(* IEC 61131-3 sources: ZPLC/conformance/cmp, 592 files *)

(* ---- cmp-042-type-from-another-file-in-a-structure-point.st ---- *)
TYPE Point : STRUCT
  x : INT;
  y : INT;
END_STRUCT END_TYPE

(* ---- cmp-042-global-in-another-file-globals.st ---- *)
VAR_GLOBAL Shared : INT; END_VAR

(* ---- cmp-042-global-initial-value-is-applied-once-globals.st ---- *)
VAR_GLOBAL
  Counter : INT := 100;
END_VAR

(* ---- cmp-042-two-tasks-share-a-global-globals.st ---- *)
VAR_GLOBAL
  Shared : INT;
END_VAR

(* ---- cmp-042-function-from-another-file-in-two-programs-lib.st ---- *)
FUNCTION Twice : INT
VAR_INPUT x : INT; END_VAR
  Twice := x * 2;
END_FUNCTION

(* ---- cmp-004-user-names-case-insensitive.st ---- *)
TYPE
  Pair : STRUCT
    Low : INT;
    High : INT;
  END_STRUCT
  Mode : (Idle, Busy);
END_TYPE

FUNCTION Twice : INT
VAR_INPUT Amount : INT; END_VAR
  TWICE := amount * 2;
END_FUNCTION

FUNCTION_BLOCK Counter
VAR_INPUT Step : INT; END_VAR
VAR_OUTPUT Total : INT; END_VAR
  total := TOTAL + step;
END_FUNCTION_BLOCK

PROGRAM Names
VAR
  P : Pair;
  C : counter;
  M : mode;
  result AT %QW0 : INT;
  is_busy AT %QX2.0 : BOOL;
END_VAR
  p.LOW := twice(AMOUNT := 3);
  p.high := TWICE(4);
  C(STEP := 5);
  c(step := 6);
  M := BUSY;
  result := P.low + p.HIGH + c.TOTAL;
  is_busy := m = busy;
END_PROGRAM

(* ---- cmp-006-missing-base-block.st ---- *)
FUNCTION_BLOCK Child EXTENDS Parent
END_FUNCTION_BLOCK

PROGRAM Caller
VAR
  c : Child;
END_VAR
END_PROGRAM

(* ---- cmp-006-property-is-rejected.st ---- *)
FUNCTION_BLOCK Holder
VAR
  stored : INT;
END_VAR
PROPERTY Value : INT
GET
  Value := stored;
END_GET
END_PROPERTY
END_FUNCTION_BLOCK

PROGRAM Props
VAR
  q AT %QW0 : INT;
END_VAR
  q := 1;
END_PROGRAM

(* ---- cmp-006-unknown-identifier-in-block-body.st ---- *)
FUNCTION_BLOCK Scale
VAR_INPUT a : INT; END_VAR
VAR_OUTPUT b : INT; END_VAR
  b := a * factor;
END_FUNCTION_BLOCK

PROGRAM Caller
VAR
  s : Scale;
  seen AT %QW0 : INT;
END_VAR
  s(a := 2);
  seen := s.b;
END_PROGRAM

(* ---- cmp-006-unknown-member-position.st ---- *)
FUNCTION_BLOCK Counter
VAR_INPUT inc : INT; END_VAR
VAR_OUTPUT total : INT; END_VAR
  total := total + inc;
END_FUNCTION_BLOCK

PROGRAM Typo
VAR
  c : Counter;
END_VAR
  c(nope := 2);
END_PROGRAM

(* ---- cmp-013-int-to-real-in-method-argument.st ---- *)
FUNCTION_BLOCK Scaler
METHOD PUBLIC Twice : REAL
VAR_INPUT
  x : REAL;
END_VAR
  Twice := x * 2.0;
END_METHOD
END_FUNCTION_BLOCK

PROGRAM Caller
VAR
  s : Scaler;
  n : INT := -3;
  r AT %QD0 : REAL;
END_VAR
  r := s.Twice(n);
END_PROGRAM

(* ---- cmp-015-interface-references-stay-one-cell-beside-64-bit-values.st ---- *)
INTERFACE IMeter
METHOD Reading : LREAL
END_METHOD
END_INTERFACE

FUNCTION_BLOCK Probe IMPLEMENTS IMeter
VAR_INPUT
  gain : LREAL;
END_VAR
METHOD Reading : LREAL
  Reading := gain + 0.5;
END_METHOD
END_FUNCTION_BLOCK

FUNCTION_BLOCK Slot
VAR_INPUT
  before : LREAL;
  meter : IMeter;
  after : LINT;
END_VAR
END_FUNCTION_BLOCK

FUNCTION Scaled : LREAL
VAR_INPUT
  source : IMeter;
  factor : LREAL;
  offset : LINT;
END_VAR
  Scaled := source.Reading() * factor + offset;
END_FUNCTION

PROGRAM WideAndInterface
VAR
  a : Probe;
  b : Probe;
  slot : Slot;
  meters : ARRAY[0..1] OF IMeter;
  wide : ARRAY[0..1] OF LINT;
  o_before AT %QD0 : LREAL;
  o_after AT %QD2 : LINT;
  o_slot AT %QD4 : LREAL;
  o_first AT %QD6 : LREAL;
  o_second AT %QD8 : LREAL;
  o_scaled AT %QD10 : LREAL;
  o_wide1 AT %QD12 : LINT;
END_VAR
  a.gain := 1.0;
  b.gain := 2.0;
  slot.before := 1.25;
  slot.meter := b;
  slot.after := -7000000000;
  meters[0] := a;
  meters[1] := b;
  wide[0] := 4294967296;
  wide[1] := -4294967296;
  o_before := slot.before;
  o_after := slot.after;
  o_slot := slot.meter.Reading();
  o_first := meters[0].Reading();
  o_second := meters[1].Reading();
  o_scaled := Scaled(meters[1], 0.1, 3000000000);
  o_wide1 := wide[1];
END_PROGRAM

(* ---- cmp-015-lreal-and-lint-keep-their-place-between-narrow-neighbours.st ---- *)
TYPE Cell :
STRUCT
  flag : BOOL;
  value : LREAL;
  tag : BYTE;
  count : LINT;
  small : INT;
END_STRUCT
END_TYPE

FUNCTION_BLOCK Holder
VAR_INPUT
  on : BOOL;
  level : LREAL;
END_VAR
VAR_OUTPUT
  seen : LINT;
  half : LREAL;
END_VAR
VAR
  steps : BYTE;
END_VAR
  steps := steps + 1;
  seen := seen + 4294967297;
  half := level / 2.0;
END_FUNCTION_BLOCK

PROGRAM WideLayout
VAR
  flag0 : BOOL;
  lone : LREAL;
  byte0 : BYTE;
  wide0 : LINT;
  int0 : INT;
  cells : ARRAY[0..2] OF Cell;
  holder : Holder;
  unit : LINT := 4294967296;
  i : DINT;
  o_flag0 AT %QX512.0 : BOOL;
  o_lone AT %QD0 : LREAL;
  o_byte0 AT %QB1024 : BYTE;
  o_wide0 AT %QD2 : LINT;
  o_int0 AT %QW600 : INT;
  o_flag1 AT %QX512.1 : BOOL;
  o_flag2 AT %QX512.2 : BOOL;
  o_value1 AT %QD4 : LREAL;
  o_value2 AT %QD6 : LREAL;
  o_tag2 AT %QB1025 : BYTE;
  o_count1 AT %QD8 : LINT;
  o_count2 AT %QD10 : LINT;
  o_small1 AT %QW601 : INT;
  o_seen AT %QD12 : LINT;
  o_half AT %QD14 : LREAL;
END_VAR
  flag0 := TRUE;
  lone := 0.1;
  byte0 := 200;
  wide0 := -4294967297;
  int0 := -3;
  FOR i := 0 TO 2 DO
    cells[i].flag := (i = 1);
    cells[i].value := 1.5 * (i + 1);
    cells[i].tag := 10 + i;
    cells[i].count := unit * (i + 1);
    cells[i].small := -100 * (i + 1);
  END_FOR;
  holder(on := TRUE, level := 0.5);
  holder(on := FALSE, level := 0.1);
  o_flag0 := flag0;
  o_lone := lone;
  o_byte0 := byte0;
  o_wide0 := wide0;
  o_int0 := int0;
  o_flag1 := cells[1].flag;
  o_flag2 := cells[2].flag;
  o_value1 := cells[1].value;
  o_value2 := cells[2].value;
  o_tag2 := cells[2].tag;
  o_count1 := cells[1].count;
  o_count2 := cells[2].count;
  o_small1 := cells[1].small;
  o_seen := holder.seen;
  o_half := holder.half;
END_PROGRAM

(* ---- cmp-015-lreal-and-lint-results-of-methods-and-interface-calls.st ---- *)
INTERFACE IMeter
METHOD Reading : LREAL
END_METHOD
METHOD Ticks : LINT
END_METHOD
END_INTERFACE

FUNCTION_BLOCK Probe IMPLEMENTS IMeter
VAR_INPUT
  gain : LREAL;
  offset : LINT;
END_VAR
METHOD Reading : LREAL
  Reading := gain * 0.1 + 0.5;
END_METHOD
METHOD Ticks : LINT
  Ticks := offset * 3;
END_METHOD
METHOD Twice : LREAL
  Twice := Reading() * 2.0;
END_METHOD
END_FUNCTION_BLOCK

FUNCTION_BLOCK FineProbe EXTENDS Probe
METHOD OVERRIDE Reading : LREAL
  Reading := SUPER^.Reading() + 0.25;
END_METHOD
METHOD OVERRIDE Ticks : LINT
  Ticks := SUPER^.Ticks() + 4294967296;
END_METHOD
END_FUNCTION_BLOCK

PROGRAM WideMethods
VAR
  plain : Probe;
  fine : FineProbe;
  meter : IMeter;
  o_reading AT %QD0 : LREAL;
  o_ticks AT %QD2 : LINT;
  o_twice AT %QD4 : LREAL;
  o_fine AT %QD6 : LREAL;
  o_fine_ticks AT %QD8 : LINT;
  o_fine_twice AT %QD10 : LREAL;
  o_through AT %QD12 : LREAL;
  o_through_ticks AT %QD14 : LINT;
  o_through_plain AT %QD16 : LREAL;
  o_after AT %QX512.0 : BOOL;
END_VAR
  plain.gain := 3.0;
  plain.offset := -2000000000;
  fine.gain := 3.0;
  fine.offset := 1;
  o_reading := plain.Reading();
  o_ticks := plain.Ticks();
  o_twice := plain.Twice();
  o_fine := fine.Reading();
  o_fine_ticks := fine.Ticks();
  o_fine_twice := fine.Twice();
  meter := fine;
  o_through := meter.Reading() + 1.0;
  o_through_ticks := meter.Ticks() - 1;
  meter := plain;
  o_through_plain := meter.Reading();
  o_after := meter.Ticks() < 0;
END_PROGRAM

(* ---- cmp-015-lreal-and-lint-through-references-and-in-out-parameters.st ---- *)
FUNCTION_BLOCK Accumulate
VAR_IN_OUT
  total : LREAL;
  count : LINT;
END_VAR
VAR_INPUT
  step : LREAL;
END_VAR
  total := total + step;
  count := count + 1;
END_FUNCTION_BLOCK

PROGRAM WideReferences
VAR
  sum : LREAL;
  big : LINT := 5000000000;
  pd : REF_TO LREAL;
  pl : REF_TO LINT;
  acc : Accumulate;
  n : LINT;
  o_sum AT %QD0 : LREAL;
  o_big AT %QD2 : LINT;
  o_count AT %QD4 : LINT;
  o_through AT %QD6 : LREAL;
END_VAR
  pd := REF(sum);
  pl := REF(big);
  acc(total := sum, count := n, step := 0.5);
  acc(total := sum, count := n, step := 0.25);
  pd^ := pd^ + 1.0;
  pl^ := pl^ * 2;
  o_sum := sum;
  o_big := big;
  o_count := n;
  o_through := pd^ * 2.0;
END_PROGRAM

(* ---- cmp-019-fb-member-int.st ---- *)
FUNCTION_BLOCK Big
VAR_OUTPUT o : INT; END_VAR
  o := 1000;
END_FUNCTION_BLOCK

PROGRAM Member
VAR
  f : Big;
  seen AT %QW0 : INT;
END_VAR
  f();
  seen := f.o;
END_PROGRAM

(* ---- cmp-019-fb-mixed-width-members.st ---- *)
FUNCTION_BLOCK Mixed
VAR_INPUT b : BYTE; END_VAR
VAR_OUTPUT i : INT; d : DINT; r : REAL; s : SINT; END_VAR
  i := -1000;
  d := -100000;
  r := 2.5;
  s := -3;
  b := 200;
END_FUNCTION_BLOCK

PROGRAM Main
VAR
  m : Mixed;
  oi AT %QW0 : INT;
  od AT %QD1 : DINT;
  orr AT %QD2 : REAL;
  os AT %QB12 : SINT;
  ob AT %QB13 : BYTE;
END_VAR
  m();
  oi := m.i;
  od := m.d;
  orr := m.r;
  os := m.s;
  ob := m.b;
END_PROGRAM

(* ---- cmp-021-fb-string-member-initial-value.st ---- *)
FUNCTION_BLOCK Named
VAR_OUTPUT label : STRING[16] := 'unit'; END_VAR
END_FUNCTION_BLOCK

PROGRAM Main
VAR
  n : Named;
  l AT %QW0 : INT;
  ok AT %QX2.0 : BOOL;
END_VAR
  n();
  l := LEN(n.label);
  ok := n.label = 'unit';
END_PROGRAM

(* ---- cmp-024-null-inside-a-function-block.st ---- *)
FUNCTION_BLOCK Probe
VAR_INPUT bind : BOOL; target : DINT; END_VAR
VAR_OUTPUT isNull : BOOL; value : DINT; END_VAR
VAR p : REF_TO DINT; END_VAR
  IF bind THEN
    p := REF(target);
  ELSE
    p := NULL;
  END_IF;
  isNull := p = NULL;
  IF NOT isNull THEN
    value := p^;
  END_IF;
END_FUNCTION_BLOCK

PROGRAM Main
VAR
  probe : Probe;
  a AT %QX0.0 : BOOL;
  b AT %QX0.1 : BOOL;
  v AT %QD1 : DINT;
END_VAR
  probe(bind := FALSE, target := 5);
  a := probe.isNull;
  probe(bind := TRUE, target := 123456);
  b := probe.isNull;
  v := probe.value;
END_PROGRAM

(* ---- cmp-025-fb-instances-keep-their-own-initial-values.st ---- *)
FUNCTION_BLOCK Start
VAR_OUTPUT v : INT := 5; END_VAR
  v := v + 1;
END_FUNCTION_BLOCK

PROGRAM Main
VAR
  f1 : Start := (v := 10);
  f2 : Start;
  a AT %QW0 : INT;
  b AT %QW1 : INT;
END_VAR
  f1();
  f2();
  a := f1.v;
  b := f2.v;
END_PROGRAM

(* ---- cmp-025-fb-member-initial-value.st ---- *)
FUNCTION_BLOCK Start
VAR_OUTPUT v : INT := 5; END_VAR
  v := v + 1;
END_FUNCTION_BLOCK

PROGRAM Members
VAR
  f : Start;
  seen AT %QW0 : INT;
END_VAR
  f();
  seen := f.v;
END_PROGRAM

(* ---- cmp-025-var-input-and-var-output-of-a-function-block.st ---- *)
FUNCTION_BLOCK Accumulate
VAR_INPUT step : INT; END_VAR
VAR_OUTPUT total : INT; END_VAR
  total := total + step;
END_FUNCTION_BLOCK

PROGRAM Inputs
VAR
  acc : Accumulate;
  result AT %QW0 : INT;
END_VAR
  acc(step := 3);
  result := acc.total;
END_PROGRAM

(* ---- cmp-026-function-block-constant-assignment-rejected.st ---- *)
FUNCTION_BLOCK Limit
VAR_OUTPUT clipped : INT; END_VAR
VAR CONSTANT MAXV : INT := 100; END_VAR
  MAXV := 5;
  clipped := MAXV;
END_FUNCTION_BLOCK

PROGRAM Main
VAR
  l : Limit;
END_VAR
  l();
END_PROGRAM

(* ---- cmp-026-function-block-constant-member.st ---- *)
FUNCTION_BLOCK Limit
VAR_INPUT v : INT; END_VAR
VAR_OUTPUT clipped : INT; END_VAR
VAR CONSTANT MAXV : INT := 100; END_VAR
  IF v > MAXV THEN
    clipped := MAXV;
  ELSE
    clipped := v;
  END_IF;
END_FUNCTION_BLOCK

PROGRAM Main
VAR
  l : Limit;
  out AT %QW0 : INT;
END_VAR
  l(v := 250);
  out := l.clipped;
END_PROGRAM

(* ---- cmp-027-fb-var-temp-initial-value-on-every-call.st ---- *)
FUNCTION_BLOCK Temp
VAR_OUTPUT o : INT; END_VAR
VAR_TEMP k : INT := 10; END_VAR
  k := k + 1;
  o := k;
END_FUNCTION_BLOCK

PROGRAM Main
VAR
  f : Temp;
  seen AT %QW0 : INT;
END_VAR
  f();
  seen := f.o;
END_PROGRAM

(* ---- cmp-027-fb-var-temp-not-retained.st ---- *)
FUNCTION_BLOCK Temp
VAR_OUTPUT o : INT; END_VAR
VAR_TEMP k : INT; END_VAR
  k := k + 1;
  o := k;
END_FUNCTION_BLOCK

PROGRAM Calls
VAR
  f : Temp;
  seen AT %QW0 : INT;
END_VAR
  f();
  seen := f.o;
END_PROGRAM

(* ---- cmp-028-in-out-bound-to-member-and-element.st ---- *)
TYPE Pt : STRUCT x : INT; z : DINT; END_STRUCT END_TYPE

FUNCTION_BLOCK Inc
VAR_IN_OUT x : INT; END_VAR
  x := x + 1;
END_FUNCTION_BLOCK

PROGRAM Main
VAR
  f : Inc;
  s : Pt;
  a : ARRAY[0..3] OF INT;
  i : INT;
  sx AT %QW0 : INT;
  a2 AT %QW1 : INT;
  a1 AT %QW2 : INT;
END_VAR
  s.x := 40;
  i := 2;
  a[2] := 7;
  f(x := s.x);
  f(x := a[i]);
  sx := s.x;
  a2 := a[2];
  a1 := a[1];
END_PROGRAM

(* ---- cmp-028-in-out-of-another-type-rejected.st ---- *)
FUNCTION_BLOCK Inc
VAR_IN_OUT x : INT; END_VAR
  x := x + 1;
END_FUNCTION_BLOCK

PROGRAM Main
VAR
  f : Inc;
  d : DINT;
END_VAR
  f(x := d);
END_PROGRAM

(* ---- cmp-028-in-out-two-instances-different-targets.st ---- *)
FUNCTION_BLOCK Inc
VAR_IN_OUT x : DINT; END_VAR
  x := x + 100000;
END_FUNCTION_BLOCK

PROGRAM Main
VAR
  f : Inc;
  g : Inc;
  a : DINT := 1;
  b : DINT := 2;
  oa AT %QD0 : DINT;
  ob AT %QD1 : DINT;
END_VAR
  f(x := a);
  g(x := b);
  f();
  oa := a;
  ob := b;
END_PROGRAM

(* ---- cmp-028-in-out-whole-structure.st ---- *)
TYPE Pt : STRUCT x : INT; z : DINT; END_STRUCT END_TYPE

FUNCTION_BLOCK Move
VAR_IN_OUT p : Pt; END_VAR
  p.x := p.x + 1;
  p.z := p.z + 100000;
END_FUNCTION_BLOCK

PROGRAM Main
VAR
  m : Move;
  point : Pt;
  ox AT %QW0 : INT;
  oz AT %QD1 : DINT;
END_VAR
  point.x := 5;
  point.z := 1;
  m(p := point);
  ox := point.x;
  oz := point.z;
END_PROGRAM

(* ---- cmp-028-unbound-in-out-faults.st ---- *)
FUNCTION_BLOCK Inc
VAR_IN_OUT x : INT; END_VAR
  x := x + 1;
END_FUNCTION_BLOCK

PROGRAM Main
VAR
  f : Inc;
END_VAR
  f();
END_PROGRAM

(* ---- cmp-028-var-in-out-by-reference.st ---- *)
FUNCTION_BLOCK Inc
VAR_IN_OUT x : INT; END_VAR
  x := x + 1;
END_FUNCTION_BLOCK

PROGRAM Reference
VAR
  f : Inc;
  v : INT := 5;
  seen AT %QW0 : INT;
END_VAR
  f(x := v);
  seen := v;
END_PROGRAM

(* ---- cmp-030-var-external-in-function-block.st ---- *)
VAR_GLOBAL
  hits : INT;
END_VAR

FUNCTION_BLOCK Counter
VAR_EXTERNAL hits : INT; END_VAR
  hits := hits + 1;
END_FUNCTION_BLOCK

PROGRAM Shared
VAR
  a : Counter;
  b : Counter;
  seen AT %QW0 : INT;
END_VAR
  a();
  b();
  seen := hits;
END_PROGRAM

(* ---- cmp-033-library-names-as-names-of-everything.st ---- *)
TYPE Reading : STRUCT Pulse : INT; Blink : INT; END_STRUCT END_TYPE

FUNCTION_BLOCK Scale
VAR_INPUT Counter : INT; END_VAR
VAR_OUTPUT Pwm : INT; END_VAR
  Pwm := Counter * 2;
END_FUNCTION_BLOCK

FUNCTION Twice : INT
VAR_INPUT Ton : INT; END_VAR
  Twice := Ton + Ton;
END_FUNCTION

PROGRAM Names
VAR
  Fifo : Reading;
  Lifo : Scale;
  Rs : INT;
  sum AT %QW0 : INT;
END_VAR
  Fifo.Pulse := 3;
  Fifo.Blink := 4;
  Lifo(Counter := Fifo.Pulse);
  Rs := Twice(Ton := Fifo.Blink);
  sum := Lifo.Pwm + Rs;
END_PROGRAM

(* ---- cmp-033-user-block-named-like-a-library-block.st ---- *)
FUNCTION_BLOCK Blink
VAR_OUTPUT level : INT; END_VAR
  level := 7;
END_FUNCTION_BLOCK

PROGRAM Own
VAR
  b : blink;
  seen AT %QW0 : INT;
END_VAR
  b();
  seen := b.level;
END_PROGRAM

(* ---- cmp-036-return-leaves-the-function-block-only.st ---- *)
FUNCTION_BLOCK Gate
VAR_INPUT go : BOOL; END_VAR
VAR_OUTPUT q : INT; END_VAR
  q := 1;
  IF go THEN
    q := 5;
    RETURN;
  END_IF;
  q := 9;
END_FUNCTION_BLOCK

PROGRAM Returns
VAR
  g : Gate;
  early AT %QW0 : INT;
  after AT %QX2.0 : BOOL;
END_VAR
  g(go := TRUE);
  early := g.q;
  after := TRUE;
END_PROGRAM

(* ---- cmp-037-output-assigned-with-colon-equals-is-rejected.st ---- *)
FUNCTION_BLOCK Adder
VAR_INPUT a : INT; END_VAR
VAR_OUTPUT sum : INT; END_VAR
  sum := a;
END_FUNCTION_BLOCK

PROGRAM Binding
VAR
  add : Adder;
END_VAR
  add(a := 1, sum := 2);
END_PROGRAM

(* ---- cmp-037-output-binding-of-a-user-block.st ---- *)
FUNCTION_BLOCK Adder
VAR_INPUT a : INT; b : INT; END_VAR
VAR_OUTPUT sum : INT; big : BOOL; END_VAR
  sum := a + b;
  big := sum > 100;
END_FUNCTION_BLOCK

PROGRAM Binding
VAR
  add : Adder;
  total AT %QW0 : INT;
  large AT %QX2.0 : BOOL;
END_VAR
  add(a := 60, b := 70, sum => total, big => large);
END_PROGRAM

(* ---- cmp-037-positional-call-of-a-user-block-is-rejected.st ---- *)
FUNCTION_BLOCK Adder
VAR_INPUT a : INT; END_VAR
VAR_OUTPUT sum : INT; END_VAR
  sum := a;
END_FUNCTION_BLOCK

PROGRAM Binding
VAR
  add : Adder;
END_VAR
  add(1);
END_PROGRAM

(* ---- cmp-037-unknown-parameter-of-a-user-block.st ---- *)
FUNCTION_BLOCK Adder
VAR_INPUT a : INT; END_VAR
VAR_OUTPUT sum : INT; END_VAR
  sum := a;
END_FUNCTION_BLOCK

PROGRAM Binding
VAR
  add : Adder;
END_VAR
  add(a := 1, nothing := 2);
END_PROGRAM

(* ---- cmp-038-array-of-user-blocks.st ---- *)
FUNCTION_BLOCK Total
VAR_INPUT inc : INT; END_VAR
VAR_OUTPUT sum : INT; END_VAR
  sum := sum + inc;
END_FUNCTION_BLOCK

PROGRAM Composition
VAR
  t : ARRAY[0..1] OF Total;
  x AT %QW0 : INT;
  y AT %QW2 : INT;
END_VAR
  t[0](inc := 1);
  t[1](inc := 10);
  x := t[0].sum;
  y := t[1].sum;
END_PROGRAM

(* ---- cmp-038-instance-inside-function-block.st ---- *)
FUNCTION_BLOCK Debounce
VAR_INPUT sig : BOOL; END_VAR
VAR_OUTPUT out : BOOL; END_VAR
VAR tmr : TON; END_VAR
  tmr(IN := sig, PT := T#20ms);
  out := tmr.Q;
END_FUNCTION_BLOCK

PROGRAM Composition
VAR
  d : Debounce;
  settled AT %QX0.0 : BOOL;
END_VAR
  d(sig := TRUE);
  settled := d.out;
END_PROGRAM

(* ---- cmp-038-timer-inside-two-instances.st ---- *)
FUNCTION_BLOCK Delay
VAR_INPUT go : BOOL; END_VAR
VAR_OUTPUT done : BOOL; END_VAR
VAR t : TON; END_VAR
  t(IN := go, PT := T#25ms);
  done := t.Q;
END_FUNCTION_BLOCK

PROGRAM Composition
VAR
  fast : Delay;
  idle : Delay;
  a AT %QX0.0 : BOOL;
  b AT %QX0.1 : BOOL;
END_VAR
  fast(go := TRUE);
  idle(go := FALSE);
  a := fast.done;
  b := idle.done;
END_PROGRAM

(* ---- cmp-038-two-instances-keep-own-state.st ---- *)
FUNCTION_BLOCK Counter
VAR_INPUT inc : INT; END_VAR
VAR_OUTPUT total : INT; END_VAR
  total := total + inc;
END_FUNCTION_BLOCK

PROGRAM Composition
VAR
  a : Counter;
  b : Counter;
  x AT %QW0 : INT;
  y AT %QW1 : INT;
END_VAR
  a(inc := 1);
  b(inc := 10);
  x := a.total;
  y := b.total;
END_PROGRAM

(* ---- cmp-039-for-inside-function-block.st ---- *)
FUNCTION_BLOCK Summer
VAR_OUTPUT s : INT; END_VAR
VAR i : INT; END_VAR
  s := 0;
  FOR i := 1 TO 4 DO
    s := s + i;
  END_FOR;
END_FUNCTION_BLOCK

PROGRAM Loop
VAR
  f : Summer;
  sum AT %QW0 : INT;
END_VAR
  f();
  sum := f.s;
END_PROGRAM

(* ---- cmp-041-abstract-block-cannot-be-instantiated.st ---- *)
FUNCTION_BLOCK ABSTRACT Template
METHOD ABSTRACT Step : INT
END_METHOD
END_FUNCTION_BLOCK

PROGRAM Abstraction
VAR
  t : Template;
END_VAR
END_PROGRAM

(* ---- cmp-041-abstract-method-is-run-by-the-derived-block.st ---- *)
FUNCTION_BLOCK ABSTRACT Template
METHOD ABSTRACT Step : INT
END_METHOD
METHOD Run : INT
  Run := Step() * 2 + 1;
END_METHOD
END_FUNCTION_BLOCK

FUNCTION_BLOCK Seven EXTENDS Template
METHOD OVERRIDE Step : INT
  Step := 7;
END_METHOD
END_FUNCTION_BLOCK

FUNCTION_BLOCK Nine EXTENDS Template
METHOD OVERRIDE Step : INT
  Step := 9;
END_METHOD
END_FUNCTION_BLOCK

PROGRAM Abstraction
VAR
  a : Seven;
  b : Nine;
  x AT %QW0 : INT;
  y AT %QW1 : INT;
END_VAR
  x := a.Run();
  y := b.Run();
END_PROGRAM

(* ---- cmp-041-abstract-method-left-unimplemented-is-rejected.st ---- *)
FUNCTION_BLOCK ABSTRACT Template
METHOD ABSTRACT Step : INT
END_METHOD
END_FUNCTION_BLOCK

FUNCTION_BLOCK Lazy EXTENDS Template
END_FUNCTION_BLOCK

PROGRAM Abstraction
VAR
  l : Lazy;
END_VAR
END_PROGRAM

(* ---- cmp-041-final-block-cannot-be-extended.st ---- *)
FUNCTION_BLOCK FINAL Sealed
END_FUNCTION_BLOCK

FUNCTION_BLOCK Open EXTENDS Sealed
END_FUNCTION_BLOCK

PROGRAM Sealing
END_PROGRAM

(* ---- cmp-041-final-method-cannot-be-overridden.st ---- *)
FUNCTION_BLOCK Base
METHOD FINAL Reading : INT
  Reading := 3;
END_METHOD
END_FUNCTION_BLOCK

FUNCTION_BLOCK Derived EXTENDS Base
METHOD OVERRIDE Reading : INT
  Reading := 4;
END_METHOD
END_FUNCTION_BLOCK

PROGRAM Derivation
VAR
  d : Derived;
  q AT %QW0 : INT;
END_VAR
  q := d.Reading();
END_PROGRAM

(* ---- cmp-041-instance-that-does-not-implement-the-interface-is-rejected.st ---- *)
INTERFACE IRun
METHOD Go : INT
END_METHOD
END_INTERFACE

FUNCTION_BLOCK Plain
METHOD Go : INT
  Go := 1;
END_METHOD
END_FUNCTION_BLOCK

PROGRAM Wrong
VAR
  p : Plain;
  r : IRun;
END_VAR
  r := p;
END_PROGRAM

(* ---- cmp-041-interface-call-of-a-null-reference-faults.st ---- *)
INTERFACE IRun
METHOD Go : INT
END_METHOD
END_INTERFACE

FUNCTION_BLOCK A IMPLEMENTS IRun
METHOD Go : INT
  Go := 1;
END_METHOD
END_FUNCTION_BLOCK

PROGRAM Unassigned
VAR
  a : A;
  r : IRun;
  seen AT %QW0 : INT;
END_VAR
  seen := 5;
  seen := r.Go();
END_PROGRAM

(* ---- cmp-041-interface-dispatch-by-the-instance-assigned.st ---- *)
INTERFACE IShape
METHOD Area : INT
END_METHOD
END_INTERFACE

FUNCTION_BLOCK Square IMPLEMENTS IShape
VAR_INPUT side : INT; END_VAR
METHOD Area : INT
  Area := side * side;
END_METHOD
END_FUNCTION_BLOCK

FUNCTION_BLOCK Rectangle IMPLEMENTS IShape
VAR_INPUT width : INT; height : INT; END_VAR
METHOD Area : INT
  Area := width * height;
END_METHOD
END_FUNCTION_BLOCK

PROGRAM Shapes
VAR
  sq : Square;
  rect : Rectangle;
  shape : IShape;
  first AT %QW0 : INT;
  second AT %QW1 : INT;
  third AT %QW2 : INT;
END_VAR
  sq.side := 4;
  rect.width := 3;
  rect.height := 5;
  shape := sq;
  first := shape.Area();
  shape := rect;
  second := shape.Area();
  sq.side := 7;
  shape := sq;
  third := shape.Area();
END_PROGRAM

(* ---- cmp-041-interface-dispatch.st ---- *)
INTERFACE IRun
METHOD Go : INT
END_METHOD
END_INTERFACE

FUNCTION_BLOCK A IMPLEMENTS IRun
METHOD Go : INT
  Go := 1;
END_METHOD
END_FUNCTION_BLOCK

PROGRAM Dispatch
VAR
  a : A;
  r : IRun;
  seen AT %QW0 : INT;
END_VAR
  r := a;
  seen := r.Go();
END_PROGRAM

(* ---- cmp-041-interface-through-inheritance-and-array-elements.st ---- *)
INTERFACE IStep
METHOD Run : INT
END_METHOD
END_INTERFACE

FUNCTION_BLOCK Base IMPLEMENTS IStep
VAR_INPUT n : INT; END_VAR
METHOD Run : INT
  Run := n;
END_METHOD
END_FUNCTION_BLOCK

FUNCTION_BLOCK Derived EXTENDS Base
METHOD OVERRIDE Run : INT
  Run := SUPER^.Run() + 1000;
END_METHOD
END_FUNCTION_BLOCK

PROGRAM Steps
VAR
  plain : ARRAY[0..2] OF Base;
  special : Derived;
  step : IStep;
  i : INT;
  total AT %QW0 : INT;
  last AT %QW1 : INT;
END_VAR
  plain[0].n := 1;
  plain[1].n := 20;
  plain[2].n := 300;
  special.n := 5;
  total := 0;
  FOR i := 0 TO 2 DO
    step := plain[i];
    total := total + step.Run();
  END_FOR;
  step := special;
  last := step.Run();
END_PROGRAM

(* ---- cmp-041-interface-variable-as-an-argument-of-a-function.st ---- *)
INTERFACE IMeasure
METHOD Read : INT
END_METHOD
END_INTERFACE

FUNCTION_BLOCK Fixed IMPLEMENTS IMeasure
METHOD Read : INT
  Read := 40;
END_METHOD
END_FUNCTION_BLOCK

FUNCTION_BLOCK Counted IMPLEMENTS IMeasure
VAR reads : INT; END_VAR
METHOD Read : INT
  reads := reads + 1;
  Read := reads;
END_METHOD
END_FUNCTION_BLOCK

FUNCTION Twice : INT
VAR_INPUT source : IMeasure; END_VAR
  Twice := source.Read() + source.Read();
END_FUNCTION

PROGRAM Sampling
VAR
  f : Fixed;
  c : Counted;
  a AT %QW0 : INT;
  b AT %QW1 : INT;
END_VAR
  a := Twice(source := f);
  b := Twice(source := c);
END_PROGRAM

(* ---- cmp-041-interface-variable-as-an-input-of-a-block.st ---- *)
INTERFACE IGain
METHOD Apply : INT
VAR_INPUT x : INT; END_VAR
END_METHOD
END_INTERFACE

FUNCTION_BLOCK Doubler IMPLEMENTS IGain
METHOD Apply : INT
VAR_INPUT x : INT; END_VAR
  Apply := x * 2;
END_METHOD
END_FUNCTION_BLOCK

FUNCTION_BLOCK Offsetter IMPLEMENTS IGain
VAR offset : INT := 100; END_VAR
METHOD Apply : INT
VAR_INPUT x : INT; END_VAR
  Apply := x + offset;
END_METHOD
END_FUNCTION_BLOCK

FUNCTION_BLOCK Stage
VAR_INPUT gain : IGain; value : INT; END_VAR
VAR_OUTPUT result : INT; END_VAR
  result := gain.Apply(value);
END_FUNCTION_BLOCK

PROGRAM Pipeline
VAR
  d : Doubler;
  o : Offsetter;
  stage : Stage;
  a AT %QW0 : INT;
  b AT %QW1 : INT;
END_VAR
  stage(gain := d, value := 21);
  a := stage.result;
  stage(gain := o, value := 21);
  b := stage.result;
END_PROGRAM

(* ---- cmp-041-method-results-of-each-type-and-inherited-statement-call.st ---- *)
FUNCTION_BLOCK Base
VAR
  n : INT;
END_VAR
METHOD Flag : BOOL
  Flag := n > 0;
END_METHOD
METHOD Small : SINT
  Small := -5;
END_METHOD
METHOD Ratio : REAL
  Ratio := 2.5;
END_METHOD
METHOD Wide : DINT
  Wide := -70000;
END_METHOD
METHOD Bump
  n := n + 1;
END_METHOD
END_FUNCTION_BLOCK

FUNCTION_BLOCK Derived EXTENDS Base
END_FUNCTION_BLOCK

PROGRAM Results
VAR
  d : Derived;
  i : INT;
  q0 AT %QX0.0 : BOOL;
  q1 AT %QB1 : SINT;
  q2 AT %QD1 : REAL;
  q3 AT %QD2 : DINT;
  q4 AT %QW6 : INT;
END_VAR
  FOR i := 1 TO 20 DO
    d.Flag();
    d.Bump();
  END_FOR;
  q0 := d.Flag();
  q1 := d.Small();
  q2 := d.Ratio();
  q3 := d.Wide();
  q4 := d.n;
END_PROGRAM

(* ---- cmp-041-method-with-several-assignments-called-in-a-loop.st ---- *)
FUNCTION_BLOCK Chooser
VAR
  calls : INT;
END_VAR
METHOD Pick : INT
VAR_INPUT
  x : INT;
END_VAR
  Pick := x;
  IF x > 5 THEN
    Pick := x * 2;
  END_IF;
  IF x > 8 THEN
    Pick := 0 - x;
  END_IF;
  calls := calls + 1;
END_METHOD
METHOD Never : INT
  calls := calls + 100;
END_METHOD
END_FUNCTION_BLOCK

PROGRAM Loop
VAR
  c : Chooser;
  i : INT;
  total : INT;
  nothing : INT := 7;
  q0 AT %QW0 : INT;
  q1 AT %QW1 : INT;
  q2 AT %QW2 : INT;
END_VAR
  total := 0;
  FOR i := 1 TO 10 DO
    total := total + c.Pick(i);
  END_FOR;
  nothing := c.Never();
  c.Pick(3);
  q0 := total;
  q1 := c.calls;
  q2 := nothing;
END_PROGRAM

(* ---- cmp-041-override-and-inherited-method.st ---- *)
FUNCTION_BLOCK Base
METHOD A : INT
  A := 1;
END_METHOD
METHOD B : INT
  B := 10;
END_METHOD
END_FUNCTION_BLOCK

FUNCTION_BLOCK Derived EXTENDS Base
METHOD OVERRIDE B : INT
  B := 20;
END_METHOD
END_FUNCTION_BLOCK

PROGRAM Inheritance
VAR
  d : Derived;
  x AT %QW0 : INT;
  y AT %QW1 : INT;
END_VAR
  x := d.A();
  y := d.B();
END_PROGRAM

(* ---- cmp-041-private-method-is-not-callable-from-a-derived-block.st ---- *)
FUNCTION_BLOCK Sensor
METHOD PRIVATE Offset : INT
  Offset := 2;
END_METHOD
END_FUNCTION_BLOCK

FUNCTION_BLOCK Scaled EXTENDS Sensor
METHOD Shifted : INT
  Shifted := Offset();
END_METHOD
END_FUNCTION_BLOCK

PROGRAM Access
VAR
  s : Scaled;
  a AT %QW0 : INT;
END_VAR
  a := s.Shifted();
END_PROGRAM

(* ---- cmp-041-private-method-is-not-callable-from-outside.st ---- *)
FUNCTION_BLOCK Gauge
METHOD PRIVATE Reading : INT
  Reading := 3;
END_METHOD
END_FUNCTION_BLOCK

PROGRAM Access
VAR
  g : Gauge;
  q AT %QW0 : INT;
END_VAR
  q := g.Reading();
END_PROGRAM

(* ---- cmp-041-protected-method-is-callable-from-a-derived-block.st ---- *)
FUNCTION_BLOCK Sensor
METHOD PROTECTED Raw : INT
  Raw := 21;
END_METHOD
METHOD PRIVATE Offset : INT
  Offset := 2;
END_METHOD
METHOD PUBLIC Corrected : INT
  Corrected := Raw() + Offset();
END_METHOD
END_FUNCTION_BLOCK

FUNCTION_BLOCK Scaled EXTENDS Sensor
METHOD Doubled : INT
  Doubled := Raw() * 2;
END_METHOD
END_FUNCTION_BLOCK

PROGRAM Access
VAR
  s : Scaled;
  a AT %QW0 : INT;
  b AT %QW1 : INT;
END_VAR
  a := s.Corrected();
  b := s.Doubled();
END_PROGRAM

(* ---- cmp-041-protected-method-is-not-callable-from-outside.st ---- *)
FUNCTION_BLOCK Gauge
METHOD PROTECTED Reading : INT
  Reading := 3;
END_METHOD
END_FUNCTION_BLOCK

PROGRAM Access
VAR
  g : Gauge;
  q AT %QW0 : INT;
END_VAR
  q := g.Reading();
END_PROGRAM

(* ---- cmp-041-public-method-is-callable.st ---- *)
FUNCTION_BLOCK Gauge
METHOD PUBLIC Reading : INT
  Reading := 3;
END_METHOD
END_FUNCTION_BLOCK

PROGRAM Access
VAR
  g : Gauge;
  q AT %QW0 : INT;
END_VAR
  q := g.Reading();
END_PROGRAM

(* ---- cmp-041-super-call-of-a-private-method-is-rejected.st ---- *)
FUNCTION_BLOCK Base
METHOD PRIVATE Secret : INT
  Secret := 1;
END_METHOD
END_FUNCTION_BLOCK

FUNCTION_BLOCK Derived EXTENDS Base
METHOD Peek : INT
  Peek := SUPER^.Secret();
END_METHOD
END_FUNCTION_BLOCK

PROGRAM P
VAR
  d : Derived;
  a AT %QW0 : INT;
END_VAR
  a := d.Peek();
END_PROGRAM

(* ---- cmp-041-super-call-runs-the-base-body.st ---- *)
FUNCTION_BLOCK Counter
VAR_OUTPUT total : INT; END_VAR
  total := total + 1;
END_FUNCTION_BLOCK

FUNCTION_BLOCK DoubleCounter EXTENDS Counter
  SUPER^();
  total := total + 10;
END_FUNCTION_BLOCK

PROGRAM Run
VAR
  c : DoubleCounter;
  seen AT %QW0 : INT;
END_VAR
  c();
  c();
  seen := c.total;
END_PROGRAM

(* ---- cmp-041-super-call-through-three-levels.st ---- *)
FUNCTION_BLOCK Base
METHOD Value : INT
  Value := 1;
END_METHOD
END_FUNCTION_BLOCK

FUNCTION_BLOCK Middle EXTENDS Base
METHOD OVERRIDE Value : INT
  Value := SUPER^.Value() + 10;
END_METHOD
END_FUNCTION_BLOCK

FUNCTION_BLOCK Top EXTENDS Middle
METHOD OVERRIDE Value : INT
  Value := SUPER^.Value() + 100;
END_METHOD
END_FUNCTION_BLOCK

PROGRAM Chain
VAR
  t : Top;
  seen AT %QW0 : INT;
END_VAR
  seen := t.Value();
END_PROGRAM

(* ---- cmp-041-super-call.st ---- *)
FUNCTION_BLOCK A
METHOD M : INT
  M := 1;
END_METHOD
END_FUNCTION_BLOCK

FUNCTION_BLOCK B EXTENDS A
METHOD OVERRIDE M : INT
  M := SUPER^.M() + 1;
END_METHOD
END_FUNCTION_BLOCK

PROGRAM Inheritance
VAR
  b : B;
  seen AT %QW0 : INT;
END_VAR
  seen := b.M();
END_PROGRAM

(* ---- cmp-041-this-member-in-method.st ---- *)
FUNCTION_BLOCK Bumper
VAR c : INT; END_VAR
METHOD Bump : INT
  THIS.c := THIS.c + 1;
  Bump := THIS.c;
END_METHOD
END_FUNCTION_BLOCK

PROGRAM Methods
VAR
  m : Bumper;
  seen AT %QW0 : INT;
END_VAR
  seen := m.Bump();
END_PROGRAM

(* ---- cmp-042-debug-map-addresses-of-every-program-lib.st ---- *)
VAR_GLOBAL
  Shared : INT;
END_VAR

FUNCTION_BLOCK Gate
VAR_INPUT open : BOOL; END_VAR
VAR_OUTPUT passed : BOOL; END_VAR
  passed := open;
END_FUNCTION_BLOCK

(* ---- cmp-042-function-block-declared-in-two-files-is-rejected-a.st ---- *)
(* the first declaration *)
FUNCTION_BLOCK Echo
END_FUNCTION_BLOCK

(* ---- cmp-042-function-block-declared-in-two-files-is-rejected-b.st ---- *)
FUNCTION_BLOCK Echo
VAR_INPUT sig : BOOL; END_VAR
END_FUNCTION_BLOCK

(* ---- cmp-042-function-block-in-another-file-echo.st ---- *)
FUNCTION_BLOCK Echo
VAR_INPUT sig : BOOL; END_VAR
VAR_OUTPUT out : BOOL; END_VAR
  out := sig;
END_FUNCTION_BLOCK

(* ---- cmp-001-undeclared-assignment-target.st ---- *)
PROGRAM Typo
VAR
  x : INT;
END_VAR
  nope := 5;
  x := 1;
END_PROGRAM

(* ---- cmp-001-undeclared-identifier-read.st ---- *)
PROGRAM Typo
VAR
  x : INT;
END_VAR
  x := nope + 1;
END_PROGRAM

(* ---- cmp-001-unknown-function.st ---- *)
PROGRAM Typo
VAR
  x : INT;
END_VAR
  x := NOSUCHFN(1);
END_PROGRAM

(* ---- cmp-002-exit-outside-loop.st ---- *)
PROGRAM Typo
VAR
  x : INT;
END_VAR
  EXIT;
  x := 1;
END_PROGRAM

(* ---- cmp-002-wrong-argument-count.st ---- *)
PROGRAM Typo
VAR
  x : INT;
END_VAR
  x := ABS();
END_PROGRAM

(* ---- cmp-003-char-is-rejected.st ---- *)
PROGRAM Character
VAR
  c : CHAR;
  q AT %QW0 : INT;
END_VAR
  q := 1;
END_PROGRAM

(* ---- cmp-003-ldate-is-rejected.st ---- *)
PROGRAM Long
VAR
  d : LDATE;
  q AT %QW0 : INT;
END_VAR
  q := 1;
END_PROGRAM

(* ---- cmp-003-ldt-is-rejected.st ---- *)
PROGRAM Long
VAR
  t : LDT;
  q AT %QW0 : INT;
END_VAR
  q := 1;
END_PROGRAM

(* ---- cmp-003-ltime-is-rejected.st ---- *)
PROGRAM Long
VAR
  t : LTIME;
  q AT %QW0 : INT;
END_VAR
  q := 1;
END_PROGRAM

(* ---- cmp-003-ltod-is-rejected.st ---- *)
PROGRAM Long
VAR
  t : LTOD;
  q AT %QW0 : INT;
END_VAR
  q := 1;
END_PROGRAM

(* ---- cmp-003-unknown-type-in-a-function-parameter.st ---- *)
FUNCTION Twice : INT
VAR_INPUT
  a : Widget;
END_VAR
  Twice := 2;
END_FUNCTION

PROGRAM Main
VAR
  x : INT;
END_VAR
  x := 1;
END_PROGRAM

(* ---- cmp-003-unknown-type-name.st ---- *)
PROGRAM Typo
VAR
  x : NoSuchType;
  y : INT;
END_VAR
  y := 1;
END_PROGRAM

(* ---- cmp-003-wchar-is-rejected.st ---- *)
PROGRAM Character
VAR
  c : WCHAR;
  q AT %QW0 : INT;
END_VAR
  q := 1;
END_PROGRAM

(* ---- cmp-004-identifier-case-insensitive.st ---- *)
PROGRAM Names
VAR
  MyVar AT %QW0 : INT;
END_VAR
  myvar := 7;
END_PROGRAM

(* ---- cmp-004-lowercase-direct-address.st ---- *)
PROGRAM Wiring
VAR
  go AT %ix0.0 : BOOL;
  lamp AT %QX0.0 : BOOL;
END_VAR
  lamp := go;
END_PROGRAM

(* ---- cmp-004-lowercase-output-member.st ---- *)
PROGRAM Timer
VAR
  t : TON;
  done AT %QX0.0 : BOOL;
END_VAR
  t(in := TRUE, pt := T#10ms);
  done := t.q;
END_PROGRAM

(* ---- cmp-004-std-block-parameter-case-insensitive.st ---- *)
PROGRAM Timer
VAR
  t : TON;
  done AT %QX0.0 : BOOL;
END_VAR
  t(in := TRUE, pt := T#10ms);
  done := t.Q;
END_PROGRAM

(* ---- cmp-004-type-name-case-insensitive.st ---- *)
program Names
var
  x : byte;
  y : int;
  seen AT %QB0 : BYTE;
end_var
  x := 5;
  y := 7;
  seen := x;
end_program

(* ---- cmp-005-bool-assigned-from-int.st ---- *)
PROGRAM Mismatch
VAR
  b : BOOL;
  i : INT;
END_VAR
  b := i + 3;
END_PROGRAM

(* ---- cmp-005-bool-assigned-to-int.st ---- *)
PROGRAM Mismatch
VAR
  b : BOOL;
  i : INT;
END_VAR
  i := b;
END_PROGRAM

(* ---- cmp-005-bool-compared-with-a-number.st ---- *)
PROGRAM Mismatch
VAR
  b : BOOL;
  i : INT;
  c : BOOL;
END_VAR
  c := b = i;
END_PROGRAM

(* ---- cmp-005-bool-in-arithmetic.st ---- *)
PROGRAM Mismatch
VAR
  b : BOOL;
  i : INT;
END_VAR
  i := i + b;
END_PROGRAM

(* ---- cmp-005-condition-is-not-a-bool.st ---- *)
PROGRAM Mismatch
VAR
  i : INT;
END_VAR
  IF i THEN i := 0; END_IF;
END_PROGRAM

(* ---- cmp-005-int-assigned-from-real.st ---- *)
PROGRAM Mismatch
VAR
  r : REAL;
  i : INT;
END_VAR
  i := r;
END_PROGRAM

(* ---- cmp-005-integer-literal-assigned-to-bool.st ---- *)
PROGRAM Mismatch
VAR
  b : BOOL;
END_VAR
  b := 1;
END_PROGRAM

(* ---- cmp-005-integer-narrowing-keeps-the-low-bits-and-warns.st ---- *)
PROGRAM Narrow
VAR
  wide : DINT := 70000;
  huge : LINT := 5000000000;
  small AT %QW0 : INT;
  low AT %QD1 : DINT;
END_VAR
  small := wide;
  low := huge;
END_PROGRAM

(* ---- cmp-005-real-assigned-to-dint.st ---- *)
PROGRAM Mismatch
VAR
  r : REAL;
  d : DINT;
END_VAR
  d := r * 2.0;
END_PROGRAM

(* ---- cmp-005-real-in-a-bit-operation.st ---- *)
PROGRAM Mismatch
VAR
  r : REAL;
  w : WORD;
END_VAR
  w := w AND r;
END_PROGRAM

(* ---- cmp-005-string-as-a-condition.st ---- *)
PROGRAM TextCondition
VAR
  text : STRING;
  n : INT;
END_VAR
  IF text THEN
    n := 1;
  END_IF;
END_PROGRAM

(* ---- cmp-005-string-as-initial-value-of-an-int.st ---- *)
PROGRAM TextInitialValue
VAR
  n : INT := 'seven';
END_VAR
END_PROGRAM

(* ---- cmp-005-string-assigned-to-bool.st ---- *)
PROGRAM TextToBool
VAR
  text : STRING;
  flag : BOOL;
END_VAR
  flag := text;
END_PROGRAM

(* ---- cmp-005-string-assigned-to-int.st ---- *)
PROGRAM TextToNumber
VAR
  text : STRING[10];
  n : INT;
END_VAR
  n := text;
END_PROGRAM

(* ---- cmp-005-string-compared-with-a-number.st ---- *)
PROGRAM TextAndNumber
VAR
  text : STRING;
  n : INT;
  same : BOOL;
END_VAR
  same := text = n;
END_PROGRAM

(* ---- cmp-005-string-length-goes-to-a-number.st ---- *)
PROGRAM Length
VAR
  text : STRING[20] := 'abcde';
  seen AT %QW0 : INT;
  where AT %QW1 : INT;
END_VAR
  seen := LEN(text);
  where := FIND(text, 'cd');
END_PROGRAM

(* ---- cmp-005-string-literal-assigned-to-time.st ---- *)
PROGRAM LiteralToTime
VAR
  t : TIME;
END_VAR
  t := 'T#1s';
END_PROGRAM

(* ---- cmp-005-string-passed-to-a-numeric-parameter.st ---- *)
FUNCTION Double : INT
VAR_INPUT
  x : INT;
END_VAR
  Double := x * 2;
END_FUNCTION

PROGRAM TextArgument
VAR
  text : STRING;
  n : INT;
END_VAR
  n := Double(x := text);
END_PROGRAM

(* ---- cmp-005-string-returned-from-a-numeric-function.st ---- *)
FUNCTION Parse : INT
VAR_INPUT
  text : STRING;
END_VAR
  Parse := text;
END_FUNCTION

PROGRAM TextReturn
VAR
  n : INT;
END_VAR
  n := Parse(text := 'x');
END_PROGRAM

(* ---- cmp-005-time-assigned-to-int.st ---- *)
PROGRAM Mismatch
VAR
  t : TIME;
  i : INT;
END_VAR
  i := t;
END_PROGRAM

(* ---- cmp-005-widening-and-explicit-conversions.st ---- *)
PROGRAM Types
VAR
  s : SINT := -3;
  u : USINT := 200;
  i : INT := 1000;
  d : DINT;
  r : REAL;
  wide AT %QD0 : DINT;
  real_out AT %QD1 : REAL;
  unsigned_out AT %QW4 : INT;
END_VAR
  d := s;
  d := d + i;
  unsigned_out := u;
  r := i;
  wide := d;
  real_out := r + 0.5;
END_PROGRAM

(* ---- cmp-005-widening-masks-and-constants-do-not-warn.st ---- *)
PROGRAM Fits
VAR
  word_value : WORD := 16#1234;
  number : DINT := 300;
  narrow : INT := 7;
  masked AT %QB0 : BYTE;
  remainder AT %QB1 : USINT;
  wider AT %QD1 : DINT;
  literal AT %QB8 : SINT;
END_VAR
  masked := word_value AND 16#FF;
  remainder := number MOD 256;
  wider := narrow;
  literal := 100 + 27;
END_PROGRAM

(* ---- cmp-005-wstring-assigned-to-real.st ---- *)
PROGRAM WideTextToReal
VAR
  text : WSTRING;
  x : REAL;
END_VAR
  x := text;
END_PROGRAM

(* ---- cmp-006-action-block-in-a-program-is-rejected.st ---- *)
PROGRAM Actions
VAR
  q AT %QW0 : INT;
END_VAR
  q := 1;

ACTION Bump
  q := q + 1;
END_ACTION
END_PROGRAM

(* ---- cmp-006-adr-is-rejected.st ---- *)
PROGRAM Addresses
VAR
  x : INT;
  p : REF_TO INT;
  q AT %QW0 : INT;
END_VAR
  p := ADR(x);
  q := 1;
END_PROGRAM

(* ---- cmp-006-array-of-arrays-is-rejected.st ---- *)
PROGRAM Nested
VAR
  a : ARRAY[1..3] OF ARRAY[1..3] OF INT;
  q AT %QW0 : INT;
END_VAR
  q := 1;
END_PROGRAM

(* ---- cmp-006-byte-order-mark.st ---- *)
PROGRAM Errors
VAR
	x : INT;
END_VAR
	x := ;
END_PROGRAM

(* ---- cmp-006-crlf-line-endings.st ---- *)
PROGRAM Errors
VAR
	x : INT;
END_VAR
	x := ;
END_PROGRAM

(* ---- cmp-006-duplicate-variable-position.st ---- *)
PROGRAM Twice
VAR
  x : INT;
  x : INT;
END_VAR
  x := 1;
END_PROGRAM

(* ---- cmp-006-enumeration-with-base-type-is-rejected.st ---- *)
TYPE Color : (Red, Green, Blue) INT; END_TYPE

PROGRAM Colours
VAR
  c : Color;
  q AT %QW0 : INT;
END_VAR
  q := 1;
END_PROGRAM

(* ---- cmp-006-namespace-is-rejected.st ---- *)
NAMESPACE Lib
FUNCTION Twice : INT
VAR_INPUT x : INT; END_VAR
  Twice := x * 2;
END_FUNCTION
END_NAMESPACE

PROGRAM Spaces
VAR
  q AT %QW0 : INT;
END_VAR
  q := 1;
END_PROGRAM

(* ---- cmp-006-operator-function-form-is-rejected.st ---- *)
PROGRAM Forms
VAR
  q AT %QW0 : INT;
END_VAR
  q := ADD(1, 2);
END_PROGRAM

(* ---- cmp-006-persistent-qualifier-is-rejected.st ---- *)
PROGRAM Kept
VAR PERSISTENT
  x : INT;
END_VAR
VAR
  q AT %QW0 : INT;
END_VAR
  q := x;
END_PROGRAM

(* ---- cmp-006-pointer-to-is-rejected.st ---- *)
PROGRAM Pointers
VAR
  x : INT;
  p : POINTER TO INT;
  q AT %QW0 : INT;
END_VAR
  q := 1;
END_PROGRAM

(* ---- cmp-006-positional-function-block-call-is-rejected.st ---- *)
PROGRAM Positional
VAR
  t : TON;
  q AT %QX0.0 : BOOL;
END_VAR
  t(TRUE, T#1s);
  q := t.Q;
END_PROGRAM

(* ---- cmp-006-subrange-type-is-rejected.st ---- *)
TYPE Percent : INT (0..100); END_TYPE

PROGRAM Ranges
VAR
  p : Percent;
  q AT %QW0 : INT;
END_VAR
  q := 1;
END_PROGRAM

(* ---- cmp-006-tab-indented-source.st ---- *)
PROGRAM Errors
VAR
	x : INT;
END_VAR
	x := ;
END_PROGRAM

(* ---- cmp-006-textual-configuration-is-rejected.st ---- *)
CONFIGURATION Plant
RESOURCE Controller ON CPU
TASK Fast(INTERVAL := T#10ms, PRIORITY := 1);
PROGRAM Main WITH Fast : Cell;
END_RESOURCE
END_CONFIGURATION

PROGRAM Cell
VAR
  q AT %QW0 : INT;
END_VAR
  q := 1;
END_PROGRAM

(* ---- cmp-006-unknown-identifier-in-function.st ---- *)
FUNCTION Half : INT
VAR_INPUT a : INT; END_VAR
  Half := a / 2;
  Half := Half + missing;
END_FUNCTION

PROGRAM Caller
VAR
  seen AT %QW0 : INT;
END_VAR
  seen := Half(4);
END_PROGRAM

(* ---- cmp-006-var-access-is-rejected.st ---- *)
VAR_ACCESS
  Reading : Shared : INT READ_ONLY;
END_VAR

PROGRAM Access
VAR
  q AT %QW0 : INT;
END_VAR
  q := 1;
END_PROGRAM

(* ---- cmp-007-declarations-and-statements.st ---- *)
PROGRAM Errors
VAR
  a : ;
  b : INT;
  c INT;
END_VAR
  b := ;
  WHILE b DO b := 1 +; END_WHILE;
END_PROGRAM

(* ---- cmp-007-lexical-and-syntax-errors.st ---- *)
PROGRAM Errors
VAR
  x : INT;
END_VAR
  x := ;
  x := 1 @ 2;
  x := 'open;
  x := ;
END_PROGRAM

(* ---- cmp-007-no-error-after-a-broken-if.st ---- *)
PROGRAM Errors
VAR
  x : INT;
END_VAR
  IF x = THEN
    x := 1;
    IF x > 1 THEN x := 2; END_IF;
  END_IF;
  x := 5;
  x := ;
END_PROGRAM

(* ---- cmp-007-three-errors-three-diagnostics.st ---- *)
PROGRAM Broken
VAR
  x : INT;
END_VAR
  x := ;
  x := 1 +;
  x := * 2;
END_PROGRAM

(* ---- cmp-007-undeclared-names-in-every-statement.st ---- *)
PROGRAM Errors
VAR
  x : INT;
END_VAR
  x := first;
  x := 1;
  x := second + 1;
  IF third THEN x := 2; END_IF;
END_PROGRAM

(* ---- cmp-008-constant-false-branch-is-not-unreachable.st ---- *)
PROGRAM Dead
VAR
  seen AT %QW0 : INT;
END_VAR
  seen := 1;
  IF FALSE THEN
    seen := 2;
  END_IF;
  seen := seen + 1;
END_PROGRAM

(* ---- cmp-008-real-literal-without-fraction-warns.st ---- *)
PROGRAM Exponent
VAR
  seen AT %QD0 : REAL;
END_VAR
  seen := 1e3;
END_PROGRAM

(* ---- cmp-008-statement-after-return-is-unreachable.st ---- *)
PROGRAM Flow
VAR
  seen AT %QW0 : INT;
END_VAR
  seen := 1;
  RETURN;
  seen := 2;
END_PROGRAM

(* ---- cmp-008-unused-variable-is-reported.st ---- *)
PROGRAM Unused
VAR
  seen AT %QW0 : INT;
  spare : INT;
END_VAR
  seen := 7;
END_PROGRAM

(* ---- cmp-008-write-only-variable-is-not-reported-by-default.st ---- *)
PROGRAM WriteOnly
VAR
  seen AT %QW0 : INT;
  scratch : INT;
END_VAR
  scratch := 3;
  seen := scratch + 1;
  scratch := 9;
END_PROGRAM

(* ---- cmp-009-block-comment-never-closed.st ---- *)
PROGRAM Open
VAR
  x : INT;
END_VAR
  x := 1;
  /* never closed
  x := 2;
END_PROGRAM

(* ---- cmp-009-comment-closed-with-the-wrong-delimiter.st ---- *)
PROGRAM Open
VAR
  x : INT;
END_VAR
  (* closed with the other kind of delimiter */
  x := 1;
END_PROGRAM

(* ---- cmp-009-error-before-an-unterminated-comment.st ---- *)
PROGRAM Open
VAR
  x : INT;
END_VAR
  x := ;
  (* never closed
END_PROGRAM

(* ---- cmp-009-parenthesis-star-comments.st ---- *)
(* A comment before the program. *)
PROGRAM Comments
VAR
  q AT %QW0 : INT;
END_VAR
  q := 1; (* a comment after a statement *)
  q := q + (* a comment inside an expression *) 2;
  (* a comment that
     spans two lines *)
  q := q * 5;
END_PROGRAM

(* ---- cmp-009-unterminated-comment-position.st ---- *)
PROGRAM Open
VAR
  x : INT;
END_VAR
  x := 1;
  (* never closed
  x := 2;
END_PROGRAM

(* ---- cmp-010-build-error-names-the-reason.st ---- *)
PROGRAM Broken
VAR
  x : INT;
END_VAR
  x := ;
END_PROGRAM

(* ---- cmp-011-abs-negative-int.st ---- *)
PROGRAM Magnitude
VAR
  value : INT := -5;
  result AT %QW0 : INT;
END_VAR
  result := ABS(value);
END_PROGRAM

(* ---- cmp-011-case-on-negative-int.st ---- *)
PROGRAM Select
VAR
  v : INT := -5;
  w : INT := -2;
  exact AT %QW0 : INT;
  ranged AT %QW2 : INT;
END_VAR
  CASE v OF
    -5: exact := 1;
    0: exact := 2;
  ELSE
    exact := 3;
  END_CASE;
  CASE w OF
    -3..-1: ranged := 10;
  ELSE
    ranged := 20;
  END_CASE;
END_PROGRAM

(* ---- cmp-011-dint-limits.st ---- *)
PROGRAM Limits
VAR
  low : DINT := -2147483648;
  high : DINT := 2147483647;
  negative AT %QX0.0 : BOOL;
  ordered AT %QX0.1 : BOOL;
  next AT %QD4 : DINT;
END_VAR
  negative := low < 0;
  ordered := high > low;
  next := low + 1;
END_PROGRAM

(* ---- cmp-011-for-loop-over-negative-int.st ---- *)
PROGRAM Count
VAR
  i : INT;
  sum AT %QW0 : INT;
  visits AT %QW2 : INT;
END_VAR
  sum := 0;
  visits := 0;
  FOR i := -3 TO 3 DO
    sum := sum + i * i * i;
    visits := visits + 1;
  END_FOR;
END_PROGRAM

(* ---- cmp-011-function-returns-negative-int.st ---- *)
FUNCTION Negate : INT
VAR_INPUT
  x : INT;
END_VAR
  Negate := 0 - x;
END_FUNCTION

PROGRAM Caller
VAR
  r AT %QW0 : INT;
  below AT %QX2.0 : BOOL;
END_VAR
  r := Negate(5);
  below := Negate(5) < 0;
END_PROGRAM

(* ---- cmp-011-int-arithmetic-positive.st ---- *)
PROGRAM Arithmetic
VAR
  a : INT := 3;
  b : INT := 4;
  c AT %QW0 : INT;
END_VAR
  c := a + b * 2;
END_PROGRAM

(* ---- cmp-011-int-compare-negative.st ---- *)
PROGRAM Compare
VAR
  level : INT := -1;
  below AT %QX0.0 : BOOL;
END_VAR
  below := level < 0;
END_PROGRAM

(* ---- cmp-011-int-direct-input.st ---- *)
PROGRAM Analog
VAR
  level AT %IW0 : INT;
  doubled AT %QW2 : INT;
  below AT %QX0.0 : BOOL;
END_VAR
  doubled := level * 2;
  below := level < 0;
END_PROGRAM

(* ---- cmp-011-int-divide-negative.st ---- *)
PROGRAM Divide
VAR
  dividend : INT := -8;
  quotient AT %QW0 : INT;
END_VAR
  quotient := dividend / 2;
END_PROGRAM

(* ---- cmp-011-int-limits.st ---- *)
PROGRAM Limits
VAR
  low : INT := -32768;
  high : INT := 32767;
  negative AT %QX0.0 : BOOL;
  ordered AT %QX0.1 : BOOL;
  span AT %QD4 : DINT;
  floor AT %QD8 : DINT;
END_VAR
  negative := low < 0;
  ordered := high > low;
  span := high - low;
  floor := low;
END_PROGRAM

(* ---- cmp-011-int-minus-one.st ---- *)
PROGRAM MinusOne
VAR
  v : INT := -1;
  negative AT %QX0.0 : BOOL;
  same AT %QX0.1 : BOOL;
  wide AT %QD4 : DINT;
END_VAR
  negative := v < 0;
  same := v = -1;
  wide := v;
END_PROGRAM

(* ---- cmp-011-int-to-real-negative.st ---- *)
PROGRAM Convert
VAR
  count : INT := -7;
  value AT %QD0 : REAL;
END_VAR
  value := INT_TO_REAL(count);
END_PROGRAM

(* ---- cmp-011-int-widens-to-dint.st ---- *)
PROGRAM Widen
VAR
  narrow : INT := -5;
  wide AT %QD0 : DINT;
END_VAR
  wide := narrow;
END_PROGRAM

(* ---- cmp-011-max-negative-int.st ---- *)
PROGRAM Largest
VAR
  low : INT := -5;
  best AT %QW0 : INT;
END_VAR
  best := MAX(low, 3);
END_PROGRAM

(* ---- cmp-011-mixed-int-dint-real.st ---- *)
PROGRAM Mixed
VAR
  small : INT := -3;
  wide : DINT := 100000;
  ratio : REAL := 0.5;
  total AT %QD0 : DINT;
  scaled AT %QD4 : REAL;
END_VAR
  total := small + wide;
  scaled := small * ratio;
END_PROGRAM

(* ---- cmp-011-sint-limits.st ---- *)
PROGRAM Limits
VAR
  low : SINT := -128;
  high : SINT := 127;
  negative AT %QX0.0 : BOOL;
  ordered AT %QX0.1 : BOOL;
  span AT %QW2 : INT;
END_VAR
  negative := low < 0;
  ordered := high > low;
  span := high - low;
END_PROGRAM

(* ---- cmp-011-sint-negative-arithmetic.st ---- *)
PROGRAM Small
VAR
  offset : SINT := -3;
  sum AT %QW0 : INT;
END_VAR
  sum := offset + 1;
END_PROGRAM

(* ---- cmp-012-literal-above-int32-as-a-dword-argument.st ---- *)
PROGRAM BigArgument
VAR
  d : DWORD := 4042322160;
  flipped AT %QD0 : DWORD;
END_VAR
  flipped := XOR_DWORD(d, 4294967295);
END_PROGRAM

(* ---- cmp-012-literal-above-int32-to-a-udint-function-parameter.st ---- *)
FUNCTION Halve : UDINT
VAR_INPUT n : UDINT; END_VAR
  Halve := n / 2;
END_FUNCTION

PROGRAM BigArgument
VAR
  out AT %QD0 : UDINT;
  typed AT %QD1 : DWORD;
END_VAR
  out := Halve(4294967294);
  typed := XOR_DWORD(DWORD#16#F0F0F0F0, 16#FFFFFFFF);
END_PROGRAM

(* ---- cmp-012-literal-above-the-range-of-a-word-parameter.st ---- *)
PROGRAM BigArgument
VAR
  w : WORD;
END_VAR
  w := AND_WORD(w, 65536);
END_PROGRAM

(* ---- cmp-012-udint-around-2-31.st ---- *)
PROGRAM Around
VAR
  below : UDINT := 2147483647;
  above : UDINT := 2147483648;
  gt AT %QX0.0 : BOOL;
  lt AT %QX0.1 : BOOL;
  ge AT %QX0.2 : BOOL;
  le AT %QX0.3 : BOOL;
END_VAR
  gt := above > below;
  lt := below < above;
  ge := above >= 2147483648;
  le := above <= below;
END_PROGRAM

(* ---- cmp-012-udint-compare-unsigned.st ---- *)
PROGRAM Big
VAR
  big : UDINT := 2147483647;
  above AT %QX0.0 : BOOL;
END_VAR
  big := big + 2000000000;
  above := big > 5;
END_PROGRAM

(* ---- cmp-012-udint-divide-and-modulo.st ---- *)
PROGRAM Divide
VAR
  a : UDINT := 4000000000;
  b : UDINT := 3000000000;
  half : UDINT := 2147483648;
  small AT %QD0 : UDINT;
  big_q AT %QD4 : UDINT;
  big_r AT %QD8 : UDINT;
  mid_q AT %QD12 : UDINT;
  mod_small AT %QD16 : UDINT;
END_VAR
  small := a / 1000;
  big_q := a / b;
  big_r := a MOD b;
  mid_q := a / half;
  mod_small := a MOD 7;
END_PROGRAM

(* ---- cmp-012-udint-divide-unsigned.st ---- *)
PROGRAM Big
VAR
  big : UDINT := 2147483647;
  third AT %QD0 : UDINT;
END_VAR
  big := big + 2000000000;
  third := big / 3;
END_PROGRAM

(* ---- cmp-012-udint-literal-above-int32.st ---- *)
PROGRAM Big
VAR
  big : UDINT := 3000000000;
  above AT %QX0.0 : BOOL;
END_VAR
  above := big > 5;
END_PROGRAM

(* ---- cmp-012-udint-max.st ---- *)
PROGRAM Largest
VAR
  top : UDINT := 4294967295;
  zero : UDINT := 0;
  gt AT %QX0.0 : BOOL;
  ge AT %QX0.1 : BOOL;
  lt AT %QX0.2 : BOOL;
  le AT %QX0.3 : BOOL;
  same AT %QX0.4 : BOOL;
END_VAR
  gt := top > zero;
  ge := top >= zero;
  lt := top < zero;
  le := top <= zero;
  same := top = 4294967295;
END_PROGRAM

(* ---- cmp-012-udint-signed-range-unchanged.st ---- *)
PROGRAM Small
VAR
  a : UDINT := 1000000;
  quotient AT %QD0 : UDINT;
  remainder AT %QD4 : UDINT;
END_VAR
  quotient := a / 7;
  remainder := a MOD 7;
END_PROGRAM

(* ---- cmp-012-udint-to-real.st ---- *)
PROGRAM Convert
VAR
  big : UDINT := 3000000000;
  r AT %QD0 : REAL;
END_VAR
  r := big;
END_PROGRAM

(* ---- cmp-012-uint-65535.st ---- *)
PROGRAM Top
VAR
  top : UINT := 65535;
  above AT %QX0.0 : BOOL;
  wide AT %QD4 : UDINT;
  wrapped AT %QW2 : UINT;
END_VAR
  above := top > 32767;
  wide := top;
  wrapped := top + 1;
END_PROGRAM

(* ---- cmp-012-uint-compare-above-int16.st ---- *)
PROGRAM Big
VAR
  big : UINT := 40000;
  above AT %QX0.0 : BOOL;
END_VAR
  above := big > 30000;
END_PROGRAM

(* ---- cmp-012-usint-holds-0-to-255.st ---- *)
PROGRAM UsintRange
VAR
  a : USINT := 200;
  b : USINT := 55;
  sum AT %QD0 : DINT;
  above AT %QX4.0 : BOOL;
  top AT %QB5 : USINT;
END_VAR
  sum := a + b;
  above := a > b;
  top := 255;
END_PROGRAM

(* ---- cmp-013-int-plus-real.st ---- *)
PROGRAM Mixed
VAR
  i : INT := -3;
  r : REAL := 0.5;
  sum AT %QD0 : REAL;
END_VAR
  sum := i + r;
END_PROGRAM

(* ---- cmp-013-int-times-real.st ---- *)
PROGRAM Scale
VAR
  count : INT := 3;
  gain : REAL := 2.0;
  scaled AT %QD0 : REAL;
END_VAR
  scaled := count * gain;
END_PROGRAM

(* ---- cmp-013-int-to-real-in-function-argument.st ---- *)
FUNCTION Twice : REAL
VAR_INPUT
  x : REAL;
END_VAR
  Twice := x * 2.0;
END_FUNCTION

PROGRAM Caller
VAR
  n : INT := -3;
  r AT %QD0 : REAL;
END_VAR
  r := Twice(n);
END_PROGRAM

(* ---- cmp-013-real-arithmetic-positive.st ---- *)
PROGRAM Arithmetic
VAR
  r : REAL := 1.5;
  q AT %QD0 : REAL;
END_VAR
  q := r * 2.0 + 0.25;
END_PROGRAM

(* ---- cmp-013-real-assigned-from-integer.st ---- *)
PROGRAM Assign
VAR
  i : INT := -4;
  init : REAL := 7;
  copy AT %QD0 : REAL;
  seven AT %QD4 : REAL;
END_VAR
  copy := i;
  seven := init;
END_PROGRAM

(* ---- cmp-013-real-compare-negative.st ---- *)
PROGRAM Order
VAR
  low : REAL;
  high : REAL;
  ordered AT %QX0.0 : BOOL;
END_VAR
  low := 0.0 - 2.0;
  high := 0.0 - 1.0;
  ordered := low < high;
END_PROGRAM

(* ---- cmp-013-real-exponent-and-boolean-literals.st ---- *)
PROGRAM Literals
VAR
  big AT %QD0 : REAL;
  small AT %QD1 : REAL;
  whole AT %QW4 : INT;
  on AT %QX10.0 : BOOL;
  off AT %QX10.1 : BOOL;
END_VAR
  big := 1.5E2;
  small := 2.5E-1;
  whole := 12345;
  on := TRUE;
  off := FALSE;
END_PROGRAM

(* ---- cmp-013-real-infinities-order.st ---- *)
PROGRAM Infinite
VAR
  bits AT %ID0 : DWORD;
  pos AT %ID0 : REAL;
  low_bits AT %ID4 : DWORD;
  neg AT %ID4 : REAL;
  big : REAL := 3.0E38;
  pos_above AT %QX0.0 : BOOL;
  neg_below AT %QX0.1 : BOOL;
  pos_same AT %QX0.2 : BOOL;
  neg_less AT %QX0.3 : BOOL;
END_VAR
  pos_above := pos > big;
  neg_below := neg < 0.0 - big;
  pos_same := pos = pos;
  neg_less := neg < pos;
END_PROGRAM

(* ---- cmp-013-real-max-min-limit-abs.st ---- *)
PROGRAM Functions
VAR
  a : REAL := -2.5;
  b : REAL := -1.5;
  hi AT %QD0 : REAL;
  lo AT %QD4 : REAL;
  clamped AT %QD8 : REAL;
  magnitude AT %QD12 : REAL;
END_VAR
  hi := MAX(a, b);
  lo := MIN(a, b);
  clamped := LIMIT(-1.0, a, 1.0);
  magnitude := ABS(a);
END_PROGRAM

(* ---- cmp-013-real-nan-is-unordered.st ---- *)
PROGRAM Unordered
VAR
  bits AT %ID0 : DWORD;
  nan AT %ID0 : REAL;
  one : REAL := 1.0;
  eq_self AT %QX0.0 : BOOL;
  ne_self AT %QX0.1 : BOOL;
  lt_one AT %QX0.2 : BOOL;
  ge_one AT %QX0.3 : BOOL;
  gt_one AT %QX0.4 : BOOL;
  le_one AT %QX0.5 : BOOL;
END_VAR
  eq_self := nan = nan;
  ne_self := nan <> nan;
  lt_one := nan < one;
  ge_one := nan >= one;
  gt_one := one > nan;
  le_one := one <= nan;
END_PROGRAM

(* ---- cmp-013-real-negate-variable.st ---- *)
PROGRAM Negate
VAR
  r : REAL := 1.5;
  q AT %QD0 : REAL;
END_VAR
  q := -r;
END_PROGRAM

(* ---- cmp-013-real-negative-literal.st ---- *)
PROGRAM Literal
VAR
  q AT %QD0 : REAL;
END_VAR
  q := -1.5;
END_PROGRAM

(* ---- cmp-013-real-negative-zero-equals-zero.st ---- *)
PROGRAM Zeros
VAR
  zero : REAL := 0.0;
  neg : REAL;
  same AT %QX0.0 : BOOL;
  below AT %QX0.1 : BOOL;
  differ AT %QX0.2 : BOOL;
END_VAR
  neg := -zero;
  same := neg = zero;
  below := neg < zero;
  differ := neg <> zero;
END_PROGRAM

(* ---- cmp-013-real-order-with-signs.st ---- *)
PROGRAM Order
VAR
  a : REAL := -2.5;
  b : REAL := -1.5;
  c : REAL := 0.0;
  d : REAL := 3.25;
  ab AT %QX0.0 : BOOL;
  bc AT %QX0.1 : BOOL;
  cd AT %QX0.2 : BOOL;
  ba AT %QX0.3 : BOOL;
  aa_le AT %QX0.4 : BOOL;
  dc_ge AT %QX0.5 : BOOL;
  ac_gt AT %QX0.6 : BOOL;
END_VAR
  ab := a < b;
  bc := b < c;
  cd := c < d;
  ba := b < a;
  aa_le := a <= a;
  dc_ge := d >= c;
  ac_gt := a > c;
END_PROGRAM

(* ---- cmp-013-real-plus-integer-literal.st ---- *)
PROGRAM Mixed
VAR
  base : REAL := 2.0;
  total AT %QD0 : REAL;
END_VAR
  total := base + 1;
END_PROGRAM

(* ---- cmp-014-and-or-xor-word.st ---- *)
PROGRAM Bits
VAR
  a : WORD := 61680;
  b : WORD := 4080;
  both AT %QW0 : WORD;
  either AT %QW2 : WORD;
  differ AT %QW4 : WORD;
END_VAR
  both := a AND b;
  either := a OR b;
  differ := a XOR b;
END_PROGRAM

(* ---- cmp-014-not-byte-in-expression.st ---- *)
PROGRAM Invert
VAR
  mask : BYTE := 15;
  above AT %QX0.0 : BOOL;
  same AT %QX0.1 : BOOL;
END_VAR
  above := (NOT mask) > 255;
  same := (NOT mask) = 240;
END_PROGRAM

(* ---- cmp-014-not-byte.st ---- *)
PROGRAM Invert
VAR
  mask : BYTE := 15;
  inverted AT %QB0 : BYTE;
END_VAR
  inverted := NOT mask;
END_PROGRAM

(* ---- cmp-014-not-dword.st ---- *)
PROGRAM Invert
VAR
  mask : DWORD := 255;
  inverted AT %QD0 : DWORD;
END_VAR
  inverted := NOT mask;
END_PROGRAM

(* ---- cmp-014-not-word.st ---- *)
PROGRAM Invert
VAR
  mask : WORD := 255;
  inverted AT %QW0 : WORD;
END_VAR
  inverted := NOT mask;
END_PROGRAM

(* ---- cmp-014-rol-byte-rotates-within-8-bits.st ---- *)
PROGRAM Rotate
VAR
  b : BYTE := 129;
  r AT %QB0 : BYTE;
  w : WORD := 32768;
  rw AT %QW2 : WORD;
END_VAR
  r := ROL(b, 1);
  rw := ROL(w, 1);
END_PROGRAM

(* ---- cmp-014-ror-word-rotates-within-16-bits.st ---- *)
PROGRAM Rotate
VAR
  w : WORD := 1;
  r AT %QW0 : WORD;
  b : BYTE := 1;
  rb AT %QB2 : BYTE;
END_VAR
  r := ROR(w, 4);
  rb := ROR(b, 1);
END_PROGRAM

(* ---- cmp-014-shl-byte-keeps-8-bits.st ---- *)
PROGRAM Shift
VAR
  b : BYTE := 200;
  past AT %QX0.0 : BOOL;
  shifted AT %QB1 : BYTE;
END_VAR
  past := SHL(b, 1) > 255;
  shifted := SHL(b, 1);
END_PROGRAM

(* ---- cmp-014-shr-and-word-logic-functions.st ---- *)
PROGRAM WordLogic
VAR
  w : WORD := 61680;
  d : DWORD := 4042322160;
  shifted AT %QW0 : WORD;
  and_w AT %QW1 : WORD;
  or_w AT %QW2 : WORD;
  xor_w AT %QW3 : WORD;
  not_w AT %QW4 : WORD;
  and_d AT %QD3 : DWORD;
  or_d AT %QD4 : DWORD;
  xor_d AT %QD5 : DWORD;
  not_d AT %QD6 : DWORD;
  ones : DWORD := 4294967295;
END_VAR
  shifted := SHR(w, 4);
  and_w := AND_WORD(w, 255);
  or_w := OR_WORD(w, 15);
  xor_w := XOR_WORD(w, 65535);
  not_w := NOT_WORD(w);
  and_d := AND_DWORD(d, 65535);
  or_d := OR_DWORD(d, 255);
  xor_d := XOR_DWORD(d, ones);
  not_d := NOT_DWORD(d);
END_PROGRAM

(* ---- cmp-015-dt-plus-time-and-difference.st ---- *)
PROGRAM Stamp
VAR
  first : DT := DT#2024-01-01-00:00:00;
  second : DT;
  later AT %QX0.0 : BOOL;
  span AT %QD1 : TIME;
END_VAR
  second := first + T#1h;
  later := second > first;
  span := second - first;
END_PROGRAM

(* ---- cmp-015-integer-width-conversion-functions.st ---- *)
PROGRAM WidthConversions
VAR
  n1 AT %QD0 : DINT;
  n2 AT %QD1 : UDINT;
  n3 AT %QW600 : INT;
  n4 AT %QB1024 : BYTE;
  w1 AT %QD2 : LINT;
  w2 AT %QD4 : LINT;
  w3 AT %QD6 : ULINT;
  w4 AT %QD8 : LWORD;
  w5 AT %QD10 : ULINT;
  w6 AT %QD12 : LINT;
  b1 AT %QX512.0 : BOOL;
  b2 AT %QX512.1 : BOOL;
  b3 AT %QX512.2 : BOOL;
  r1 AT %QD14 : LREAL;
END_VAR
  n1 := LINT_TO_DINT(5000000000);
  n2 := ULINT_TO_UDINT(18446744073709551615);
  n3 := LINT_TO_INT(-4294967297);
  n4 := LWORD_TO_BYTE(16#1234567890ABCDEF);
  w1 := DINT_TO_LINT(-1);
  w2 := UDINT_TO_LINT(4294967295);
  w3 := DINT_TO_ULINT(-1);
  w4 := BYTE_TO_LWORD(200);
  w5 := LINT_TO_ULINT(-1);
  w6 := ULINT_TO_LINT(18446744073709551615);
  b1 := LINT_TO_BOOL(0);
  b2 := LINT_TO_BOOL(4294967296);
  b3 := LWORD_TO_BOOL(16#8000000000000000);
  r1 := LINT_TO_LREAL(-1);
END_PROGRAM

(* ---- cmp-015-lint-abs-and-negate.st ---- *)
PROGRAM AbsNeg
VAR
  neg : LINT := -9000000000;
  min : LINT := -9223372036854775808;
  pos : LINT := 9000000000;
  a1 AT %QD0 : LINT;
  a2 AT %QD2 : LINT;
  a3 AT %QD4 : LINT;
  n1 AT %QD6 : LINT;
  n2 AT %QD8 : LINT;
  n3 AT %QD10 : LINT;
END_VAR
  a1 := ABS(neg);
  a2 := ABS(min);
  a3 := ABS(pos);
  n1 := -neg;
  n2 := -min;
  n3 := -pos;
END_PROGRAM

(* ---- cmp-015-lint-add-and-subtract-carry.st ---- *)
PROGRAM Carry
VAR
  a : LINT := 4294967295;
  up : LINT;
  down : LINT;
  zero : LINT := 0;
  one : LINT := 1;
  below : LINT;
  carried AT %QX0.0 : BOOL;
  borrowed AT %QX0.1 : BOOL;
  negative AT %QX0.2 : BOOL;
  back AT %QX0.3 : BOOL;
END_VAR
  up := a + 1;
  down := up - 1;
  below := zero - one;
  carried := up = 4294967296;
  borrowed := down = 4294967295;
  negative := below < 0;
  back := below + one = 0;
END_PROGRAM

(* ---- cmp-015-lint-and-lword-bit-access.st ---- *)
PROGRAM WideBits
VAR
  w : LWORD := 16#0000000100000000;
  l : LINT;
  b32 AT %QX512.0 : BOOL;
  b31 AT %QX512.1 : BOOL;
  o_l AT %QD0 : LINT;
  o_w AT %QD2 : LWORD;
END_VAR
  b32 := w.32;
  b31 := w.31;
  l := 0;
  l.63 := TRUE;
  l.0 := TRUE;
  w.63 := TRUE;
  w.32 := FALSE;
  o_l := l;
  o_w := w;
END_PROGRAM

(* ---- cmp-015-lint-case-selector-and-labels.st ---- *)
PROGRAM WideCase
VAR
  sel : LINT;
  r1 AT %QD0 : DINT;
  r2 AT %QD1 : DINT;
  r3 AT %QD2 : DINT;
  r4 AT %QD3 : DINT;
END_VAR
  sel := 5000000000;
  CASE sel OF
    1: r1 := 1;
    5000000000: r1 := 2;
    -5000000000: r1 := 3;
  ELSE r1 := 9;
  END_CASE;
  sel := -5000000000;
  CASE sel OF
    1: r2 := 1;
    5000000000: r2 := 2;
    -5000000000: r2 := 3;
  ELSE r2 := 9;
  END_CASE;
  sel := 9000000000000000000;
  CASE sel OF
    1..10: r3 := 1;
    8000000000000000000..9223372036854775807: r3 := 2;
  ELSE r3 := 9;
  END_CASE;
  sel := 77;
  CASE sel OF
    1..10: r4 := 1;
    4294967296: r4 := 2;
  END_CASE;
  r4 := r4 + 40;
END_PROGRAM

(* ---- cmp-015-lint-compare-signed-and-unsigned-order.st ---- *)
PROGRAM Order
VAR
  sl : LINT := -1;
  su : ULINT := 18446744073709551615;
  zero : LINT := 0;
  zu : ULINT := 0;
  lo : LINT := -9223372036854775808;
  hi : LINT := 9223372036854775807;
  w1 : LWORD := 16#8000000000000000;
  w2 : LWORD := 16#7FFFFFFFFFFFFFFF;
  a AT %QX512.0 : BOOL;
  b AT %QX512.1 : BOOL;
  c AT %QX512.2 : BOOL;
  d AT %QX512.3 : BOOL;
  e AT %QX512.4 : BOOL;
  f AT %QX512.5 : BOOL;
  g AT %QX512.6 : BOOL;
  h AT %QX512.7 : BOOL;
  i AT %QX513.0 : BOOL;
  j AT %QX513.1 : BOOL;
  k AT %QX513.2 : BOOL;
END_VAR
  a := sl < zero;
  b := su > zu;
  c := lo < hi;
  d := lo <= lo;
  e := hi >= hi;
  f := w1 > w2;
  g := w1 = 16#8000000000000000;
  h := sl <> zero;
  i := hi > lo;
  j := su < zu;
  k := (lo + hi) = -1;
END_PROGRAM

(* ---- cmp-015-lint-division-by-zero-faults.st ---- *)
PROGRAM ByZero
VAR
  n : LINT := 5;
  z : LINT;
  r AT %QD0 : LINT;
END_VAR
  r := n / z;
END_PROGRAM

(* ---- cmp-015-lint-division-truncates-toward-zero.st ---- *)
PROGRAM Quotients
VAR
  p7 : LINT := 7;
  m7 : LINT := -7;
  p2 : LINT := 2;
  m2 : LINT := -2;
  p3 : LINT := 3;
  m3 : LINT := -3;
  big : LINT := 1000000000000;
  seven : LINT := 7;
  min : LINT := -9223372036854775808;
  m1 : LINT := -1;
  max : LINT := 9223372036854775807;
  q1 AT %QD0 : LINT;
  q2 AT %QD2 : LINT;
  q3 AT %QD4 : LINT;
  q4 AT %QD6 : LINT;
  q5 AT %QD8 : LINT;
  q6 AT %QD10 : LINT;
  q7 AT %QD12 : LINT;
  r1 AT %QD14 : LINT;
  r2 AT %QD16 : LINT;
  r3 AT %QD18 : LINT;
  r4 AT %QD20 : LINT;
  r5 AT %QD22 : LINT;
  r6 AT %QD24 : LINT;
END_VAR
  q1 := p7 / p2;
  q2 := m7 / p2;
  q3 := p7 / m2;
  q4 := m7 / m2;
  q5 := big / seven;
  q6 := min / m1;
  q7 := max / m1;
  r1 := p7 MOD p3;
  r2 := m7 MOD p3;
  r3 := p7 MOD m3;
  r4 := big MOD seven;
  r5 := min MOD m1;
  r6 := m7 MOD m3;
END_PROGRAM

(* ---- cmp-015-lint-extreme-values.st ---- *)
PROGRAM Extremes
VAR
  top : LINT := 9223372036854775807;
  bottom : LINT := -9223372036854775808;
  ordered AT %QX0.0 : BOOL;
  sum AT %QX0.1 : BOOL;
  wraps AT %QX0.2 : BOOL;
  negated AT %QX0.3 : BOOL;
END_VAR
  ordered := top > bottom;
  sum := top + bottom = -1;
  wraps := top + 1 = bottom;
  negated := -top = bottom + 1;
END_PROGRAM

(* ---- cmp-015-lint-for-counter-crosses-32-bits.st ---- *)
PROGRAM WideFor
VAR
  i : LINT;
  sum : LINT;
  n : LINT;
  down : LINT;
  res_sum AT %QD0 : LINT;
  res_n AT %QD2 : LINT;
  res_down AT %QD4 : LINT;
  res_i AT %QD6 : LINT;
END_VAR
  sum := 0;
  FOR i := 4294967294 TO 4294967298 DO
    sum := sum + i;
    n := n + 1;
  END_FOR;
  down := 0;
  FOR i := 4294967298 TO 4294967294 BY -2 DO
    down := down + 1;
  END_FOR;
  res_sum := sum;
  res_n := n;
  res_down := down;
  res_i := i;
END_PROGRAM

(* ---- cmp-015-lint-function-parameter-and-result.st ---- *)
FUNCTION AddOne : LINT
VAR_INPUT
  x : LINT;
END_VAR
  AddOne := x + 1;
END_FUNCTION

PROGRAM Caller
VAR
  start : LINT := 4294967295;
  r : LINT;
  ok AT %QX0.0 : BOOL;
END_VAR
  r := AddOne(start);
  ok := r = 4294967296;
END_PROGRAM

(* ---- cmp-015-lint-literal-above-int32.st ---- *)
PROGRAM Wide
VAR
  big : LINT := 5000000000;
  above AT %QX0.0 : BOOL;
END_VAR
  above := big > 4294967296;
END_PROGRAM

(* ---- cmp-015-lint-literals-over-the-full-range.st ---- *)
PROGRAM Literals
VAR
  a : LINT := -9223372036854775808;
  b : LINT := 9223372036854775807;
  c : ULINT := 18446744073709551615;
  d : LWORD := 16#FFFFFFFFFFFFFFFF;
  e : LWORD := 16#DEADBEEFCAFEBABE;
  f : LINT := 16#7FFFFFFFFFFFFFFF;
  g : ULINT := 8#1777777777777777777777;
  h : LWORD := 2#1000000000000000000000000000000000000000000000000000000000000001;
  i : LINT := LINT#-9;
  j : LWORD := LWORD#16#FF00;
  k : LREAL := LREAL#0.1;
  o_a AT %QD0 : LINT;
  o_b AT %QD2 : LINT;
  o_f AT %QD4 : LINT;
  o_c AT %QD6 : ULINT;
  o_d AT %QD8 : LWORD;
  o_e AT %QD10 : LWORD;
  o_g AT %QD12 : ULINT;
  o_h AT %QD14 : LWORD;
  o_i AT %QD16 : LINT;
  o_j AT %QD18 : LWORD;
  o_k AT %QD20 : LREAL;
  o_typed AT %QD22 : LINT;
END_VAR
  o_a := a;
  o_b := b;
  o_f := f;
  o_c := c;
  o_d := d;
  o_e := e;
  o_g := g;
  o_h := h;
  o_i := i;
  o_j := j;
  o_k := k;
  o_typed := LINT#4294967296 + LINT#1;
END_PROGRAM

(* ---- cmp-015-lint-mixed-width-arithmetic.st ---- *)
PROGRAM Mixed
VAR
  small : DINT := -2147483648;
  unsigned : UDINT := 4294967295;
  wide : LINT := 1000000;
  s1 AT %QD0 : LINT;
  s2 AT %QD2 : LINT;
  s3 AT %QD4 : LINT;
  s4 AT %QD6 : LINT;
  s5 AT %QD8 : LINT;
  gt AT %QX512.0 : BOOL;
  ge_unsigned AT %QX512.1 : BOOL;
END_VAR
  s1 := wide * small;
  s2 := wide + unsigned;
  s3 := small - wide;
  s4 := wide * 4000000000;
  s5 := wide / small;
  gt := wide > small;
  ge_unsigned := wide * 5000 >= unsigned;
END_PROGRAM

(* ---- cmp-015-lint-modulo-by-zero-faults.st ---- *)
PROGRAM ByZero
VAR
  n : LINT := 5;
  z : LINT;
  r AT %QD0 : LINT;
END_VAR
  r := n MOD z;
END_PROGRAM

(* ---- cmp-015-lint-multiplication-wraps-at-64-bits.st ---- *)
PROGRAM Product
VAR
  a : LINT := 3;
  b : LINT := 4;
  c : LINT := 4294967295;
  d : LINT := -3;
  e : LINT := 4294967296;
  f : LINT := 9223372036854775807;
  g : LINT := -9223372036854775808;
  h : LINT := -1;
  i : LINT := 123456789012;
  j : LINT := 987;
  p1 AT %QD0 : LINT;
  p2 AT %QD2 : LINT;
  p3 AT %QD4 : LINT;
  p4 AT %QD6 : LINT;
  p5 AT %QD8 : LINT;
  p6 AT %QD10 : LINT;
  p7 AT %QD12 : LINT;
  p8 AT %QD14 : LINT;
END_VAR
  p1 := a * b;
  p2 := c * c;
  p3 := d * b;
  p4 := e * e;
  p5 := f * 2;
  p6 := g * h;
  p7 := i * j;
  p8 := -e * e;
END_PROGRAM

(* ---- cmp-015-lint-small-value.st ---- *)
PROGRAM Wide
VAR
  count : LINT := 5;
  ok AT %QX0.0 : BOOL;
END_VAR
  count := count + 1;
  ok := count = 6;
END_PROGRAM

(* ---- cmp-015-lint-widens-and-narrows.st ---- *)
PROGRAM Convert
VAR
  signed : DINT := -5;
  unsigned : UDINT := 4294967295;
  from_signed : LINT;
  from_unsigned : LINT;
  wide : LINT := 5000000000;
  low AT %QD1 : DINT;
  same AT %QX0.0 : BOOL;
  positive AT %QX0.1 : BOOL;
END_VAR
  from_signed := signed;
  from_unsigned := unsigned;
  low := wide;
  same := from_signed = -5;
  positive := from_unsigned = 4294967295;
END_PROGRAM

(* ---- cmp-015-lreal-abs-sqrt-limit-select.st ---- *)
PROGRAM DoubleFunctions
VAR
  a : LREAL := -2.0;
  two : LREAL := 2.0;
  neg : LREAL := -4.0;
  tiny : LREAL := 1.0E-310;
  lo : LREAL := -1.5;
  hi : LREAL := 1.5;
  x : LREAL := 7.25;
  la : LINT := -5000000000;
  lb : LINT := 6000000000;
  sel : BOOL := TRUE;
  k : DINT := 2;
  f1 AT %QD0 : LREAL;
  f2 AT %QD2 : LREAL;
  f3 AT %QD4 : LREAL;
  f4 AT %QD6 : LREAL;
  f5 AT %QD8 : LREAL;
  f6 AT %QD10 : LREAL;
  f7 AT %QD12 : LREAL;
  f8 AT %QD14 : LREAL;
  f9 AT %QD16 : LREAL;
  f10 AT %QD18 : LREAL;
  f11 AT %QD20 : LREAL;
  g1 AT %QD22 : LINT;
  g2 AT %QD24 : LINT;
  g3 AT %QD26 : LINT;
  g4 AT %QD28 : LINT;
  g5 AT %QD30 : LINT;
  g6 AT %QD32 : LINT;
END_VAR
  f1 := ABS(a);
  f2 := SQRT(two);
  f3 := SQRT(neg);
  f4 := SQRT(tiny);
  f5 := MAX(a, two);
  f6 := MIN(a, two);
  f7 := LIMIT(lo, x, hi);
  f8 := LIMIT(lo, -9.0, hi);
  f9 := LIMIT(lo, 0.25, hi);
  f10 := SEL(sel, a, two);
  f11 := MUX(k, a, two, x);
  g1 := MAX(la, lb);
  g2 := MIN(la, lb);
  g3 := LIMIT(-1000000000000, la, 1000000000000);
  g4 := LIMIT(0, la, lb);
  g5 := SEL(sel, la, lb);
  g6 := MUX(0, la, lb);
END_PROGRAM

(* ---- cmp-015-lreal-addition-subtraction-keep-52-bits.st ---- *)
PROGRAM DoubleSum
VAR
  a : LREAL := 0.1;
  b : LREAL := 0.2;
  big : LREAL := 10000000000.0;
  huge : LREAL := 1.0E16;
  tiny : LREAL := 1.0E-300;
  s1 AT %QD0 : LREAL;
  s2 AT %QD2 : LREAL;
  s3 AT %QD4 : LREAL;
  s4 AT %QD6 : LREAL;
  s5 AT %QD8 : LREAL;
  s6 AT %QD10 : LREAL;
  s7 AT %QD12 : LREAL;
  s8 AT %QD14 : LREAL;
END_VAR
  s1 := a + b;
  s2 := b - a;
  s3 := big + 1.0;
  s4 := huge + 1.0;
  s5 := huge + 3.0;
  s6 := tiny + huge;
  s7 := a - a;
  s8 := -a - b;
END_PROGRAM

(* ---- cmp-015-lreal-and-lint-globals-members-and-retained-start-from-their-initial-values.st ---- *)
TYPE Reading :
STRUCT
  weight : LREAL := 0.1;
  count : LINT := -5000000000;
  tag : INT := 7;
END_STRUCT
END_TYPE

VAR_GLOBAL
  g_double : LREAL := 0.1;
  g_wide : LINT := 5000000000;
  g_top : ULINT := 18446744073709551615;
  g_row : ARRAY[0..2] OF LREAL := [1.5, 2.5, 3.5];
  g_reading : Reading;
END_VAR

VAR_GLOBAL RETAIN
  g_kept : LREAL := 100.25;
  g_hits : LINT := 4294967296;
END_VAR

PROGRAM WideInitial
VAR
  o_double AT %QD0 : LREAL;
  o_wide AT %QD2 : LINT;
  o_top AT %QD4 : ULINT;
  o_row2 AT %QD6 : LREAL;
  o_weight AT %QD8 : LREAL;
  o_count AT %QD10 : LINT;
  o_tag AT %QW600 : INT;
  o_kept AT %QD12 : LREAL;
  o_hits AT %QD14 : LINT;
END_VAR
  g_kept := g_kept * 2.0;
  g_hits := g_hits + 1;
  o_double := g_double;
  o_wide := g_wide;
  o_top := g_top;
  o_row2 := g_row[2];
  o_weight := g_reading.weight;
  o_count := g_reading.count;
  o_tag := g_reading.tag;
  o_kept := g_kept;
  o_hits := g_hits;
END_PROGRAM

(* ---- cmp-015-lreal-and-lint-in-arrays-structures-and-calls.st ---- *)
TYPE Sample :
STRUCT
  weight : LREAL;
  count : LINT;
  flag : BOOL;
END_STRUCT
END_TYPE

FUNCTION Lerp : LREAL
VAR_INPUT
  a : LREAL;
  b : LREAL;
  t : LREAL;
END_VAR
  Lerp := a + (b - a) * t;
END_FUNCTION

FUNCTION Scale : LINT
VAR_INPUT
  base : LINT;
  factor : ULINT;
END_VAR
  Scale := base * factor;
END_FUNCTION

PROGRAM WidePlaces
VAR
  values : ARRAY[0..3] OF LREAL := [0.5, 0.25, 0.125, 0.0625];
  counts : ARRAY[1..3] OF LINT := [10000000000, -20000000000, 30000000000];
  s : Sample;
  sum : LREAL;
  total : LINT;
  i : DINT;
  o_sum AT %QD0 : LREAL;
  o_total AT %QD2 : LINT;
  o_weight AT %QD4 : LREAL;
  o_count AT %QD6 : LINT;
  o_flag AT %QX512.0 : BOOL;
  o_lerp AT %QD8 : LREAL;
  o_lerp2 AT %QD10 : LREAL;
  o_scale AT %QD12 : LINT;
END_VAR
  sum := 0.0;
  total := 0;
  FOR i := 0 TO 3 DO
    sum := sum + values[i];
  END_FOR;
  FOR i := 1 TO 3 DO
    total := total + counts[i];
  END_FOR;
  s.weight := 0.1;
  s.count := 5000000000;
  s.flag := TRUE;
  s.weight := s.weight + 0.2;
  s.count := s.count * 3;
  o_sum := sum;
  o_total := total;
  o_weight := s.weight;
  o_count := s.count;
  o_flag := s.flag;
  o_lerp := Lerp(1.0, 2.0, 0.1);
  o_lerp2 := Lerp(values[0], values[3], 0.5);
  o_scale := Scale(-3000000000, 4);
END_PROGRAM

(* ---- cmp-015-lreal-comparisons-and-nan.st ---- *)
PROGRAM DoubleCompare
VAR
  one : LREAL := 1.0;
  two : LREAL := 2.0;
  nzero : LREAL := -0.0;
  zero : LREAL := 0.0;
  max : LREAL := 1.7976931348623157E308;
  inf : LREAL;
  nan : LREAL;
  close : LREAL := 1.0000000000000002;
  lt AT %QX512.0 : BOOL;
  le AT %QX512.1 : BOOL;
  gt AT %QX512.2 : BOOL;
  ge AT %QX512.3 : BOOL;
  eq0 AT %QX512.4 : BOOL;
  lt0 AT %QX512.5 : BOOL;
  ne_close AT %QX512.6 : BOOL;
  lt_close AT %QX512.7 : BOOL;
  inf_gt AT %QX513.0 : BOOL;
  neg_inf_lt AT %QX513.1 : BOOL;
  nan_eq AT %QX513.2 : BOOL;
  nan_ne AT %QX513.3 : BOOL;
  nan_lt AT %QX513.4 : BOOL;
  nan_gt AT %QX513.5 : BOOL;
  nan_le AT %QX513.6 : BOOL;
  nan_ge AT %QX513.7 : BOOL;
  inf_eq AT %QX514.0 : BOOL;
END_VAR
  inf := max * 10.0;
  nan := inf - inf;
  lt := one < two;
  le := one <= one;
  gt := two > one;
  ge := two >= two;
  eq0 := nzero = zero;
  lt0 := nzero < zero;
  ne_close := one <> close;
  lt_close := one < close;
  inf_gt := inf > max;
  neg_inf_lt := -inf < -max;
  nan_eq := nan = nan;
  nan_ne := nan <> nan;
  nan_lt := nan < one;
  nan_gt := nan > one;
  nan_le := one <= nan;
  nan_ge := nan >= nan;
  inf_eq := inf = inf;
END_PROGRAM

(* ---- cmp-015-lreal-conversion-functions.st ---- *)
PROGRAM DoubleConversions
VAR
  h : LREAL := 2.5;
  h3 : LREAL := 3.5;
  n : LREAL := -2.5;
  big : LREAL := 1.0E30;
  neg : LREAL := -1.0E30;
  exact : LREAL := 9007199254740992.0;
  three : LREAL := 3.9;
  zero : LREAL := 0.0;
  nan : LREAL;
  rbig : REAL := 16777216.0;
  d1 AT %QD0 : DINT;
  d2 AT %QD1 : DINT;
  d3 AT %QD2 : DINT;
  d4 AT %QD3 : DINT;
  d5 AT %QD4 : DINT;
  d6 AT %QD5 : DINT;
  d7 AT %QD6 : DINT;
  u1 AT %QD7 : UDINT;
  u2 AT %QD8 : UDINT;
  u3 AT %QD9 : UDINT;
  s1 AT %QB1024 : SINT;
  l1 AT %QD10 : LINT;
  l2 AT %QD12 : LINT;
  l3 AT %QD14 : LINT;
  l4 AT %QD16 : LINT;
  l5 AT %QD18 : ULINT;
  l6 AT %QD20 : ULINT;
  l7 AT %QD22 : ULINT;
  f1 AT %QD24 : REAL;
  e1 AT %QD25 : LREAL;
  e2 AT %QD27 : LREAL;
  e3 AT %QD29 : LREAL;
  e4 AT %QD31 : LREAL;
  e5 AT %QD33 : LREAL;
  e6 AT %QD35 : LREAL;
  b1 AT %QX512.0 : BOOL;
  b2 AT %QX512.1 : BOOL;
  b3 AT %QX512.2 : BOOL;
  f2 AT %QD37 : REAL;
  f3 AT %QD38 : REAL;
END_VAR
  nan := (1.0E308 * 10.0) - (1.0E308 * 10.0);
  d1 := LREAL_TO_DINT(h);
  d2 := LREAL_TO_DINT(h3);
  d3 := LREAL_TO_DINT(n);
  d4 := LREAL_TO_DINT(big);
  d5 := LREAL_TO_DINT(neg);
  d6 := LREAL_TO_DINT(nan);
  d7 := LREAL_TO_DINT(three);
  u1 := LREAL_TO_UDINT(big);
  u2 := LREAL_TO_UDINT(n);
  u3 := LREAL_TO_UDINT(3000000000.4);
  s1 := LREAL_TO_SINT(300.0);
  l1 := LREAL_TO_LINT(exact);
  l2 := LREAL_TO_LINT(neg);
  l3 := LREAL_TO_LINT(big);
  l4 := LREAL_TO_LINT(n);
  l5 := LREAL_TO_ULINT(big);
  l6 := LREAL_TO_ULINT(n);
  l7 := LREAL_TO_ULINT(18446744073709549568.0);
  f1 := LREAL_TO_REAL(0.1);
  e1 := REAL_TO_LREAL(rbig);
  e2 := LINT_TO_LREAL(-9007199254740993);
  e3 := ULINT_TO_LREAL(18446744073709551615);
  e4 := DINT_TO_LREAL(-5);
  e5 := UDINT_TO_LREAL(4294967295);
  e6 := LWORD_TO_LREAL(16#8000000000000000);
  b1 := LREAL_TO_BOOL(zero);
  b2 := LREAL_TO_BOOL(h);
  b3 := LREAL_TO_BOOL(nan);
  f2 := LINT_TO_REAL(1152921573326323713);
  f3 := ULINT_TO_REAL(18446744073709551615);
END_PROGRAM

(* ---- cmp-015-lreal-division-by-zero-faults.st ---- *)
PROGRAM DoubleByZero
VAR
  n : LREAL := 1.0;
  z : LREAL;
  r AT %QD0 : LREAL;
END_VAR
  r := n / z;
END_PROGRAM

(* ---- cmp-015-lreal-double-precision.st ---- *)
PROGRAM Precise
VAR
  x : LREAL := 10000000000.0;
  grew AT %QX0.0 : BOOL;
END_VAR
  x := x + 1.0;
  grew := x > 10000000000.0;
END_PROGRAM

(* ---- cmp-015-lreal-keeps-its-value-between-scans.st ---- *)
PROGRAM Accumulate
VAR
  acc : LREAL;
  n : LINT := 4294967295;
  o_acc AT %QD0 : LREAL;
  o_n AT %QD2 : LINT;
  o_kept AT %QD4 : LREAL;
END_VAR
VAR RETAIN
  kept : LREAL := 100.25;
END_VAR
  acc := acc + 0.1;
  n := n + 1;
  kept := kept * 2.0;
  o_acc := acc;
  o_n := n;
  o_kept := kept;
END_PROGRAM

(* ---- cmp-015-lreal-literal-takes-the-type-of-its-context.st ---- *)
VAR_GLOBAL CONSTANT
  PI_REAL : REAL := 3.14159;
  PI_LREAL : LREAL := 3.14159;
  SIZE : DINT := 7;
END_VAR

PROGRAM DoubleContext
VAR
  x : LREAL := 0.0;
  half : LREAL := 0.5;
  c1 AT %QD0 : LREAL;
  c2 AT %QD2 : LREAL;
  c3 AT %QD4 : LREAL;
  c4 AT %QD6 : LREAL;
  c5 AT %QD8 : LREAL;
  c6 AT %QD10 : LREAL;
  c7 AT %QD12 : LREAL;
  k1 AT %QD14 : LREAL;
  k2 AT %QD16 : LREAL;
  k3 AT %QD18 : LREAL;
END_VAR
  c1 := 0.1 + 0.2;
  c2 := x + 0.1;
  c3 := half * 0.1;
  c4 := REAL#0.1 + x;
  c5 := LREAL#0.1 * 3;
  c6 := 1.0 / 3.0;
  c7 := -0.5 * 4;
  k1 := PI_REAL * 2.0;
  k2 := PI_LREAL * 2.0;
  k3 := SIZE / 2 + 0.5;
END_PROGRAM

(* ---- cmp-015-lreal-literals-with-exponent.st ---- *)
PROGRAM DoubleLiterals
VAR
  a : LREAL := 1.0E-3;
  b : LREAL := 1.5E2;
  c : LREAL := 2.5e-3;
  d : LREAL := 1.7976931348623157E308;
  e : LREAL := 4.9E-324;
  f : LREAL := -123456789.123456789;
  g : LREAL := 3.141592653589793;
  h : LREAL := 100;
  i : LREAL := -7;
  j : LREAL := 1.0E+10;
  o_a AT %QD0 : LREAL;
  o_b AT %QD2 : LREAL;
  o_c AT %QD4 : LREAL;
  o_d AT %QD6 : LREAL;
  o_e AT %QD8 : LREAL;
  o_f AT %QD10 : LREAL;
  o_g AT %QD12 : LREAL;
  o_h AT %QD14 : LREAL;
  o_i AT %QD16 : LREAL;
  o_j AT %QD18 : LREAL;
END_VAR
  o_a := a;
  o_b := b;
  o_c := c;
  o_d := d;
  o_e := e;
  o_f := f;
  o_g := g;
  o_h := h;
  o_i := i;
  o_j := j;
END_PROGRAM

(* ---- cmp-015-lreal-mixed-with-integers-and-real.st ---- *)
PROGRAM DoubleMixed
VAR
  d : LREAL := 0.5;
  i : DINT := -3;
  u : UDINT := 4294967295;
  l : LINT := 9007199254740993;
  r : REAL := 0.1;
  w : ULINT := 18446744073709551615;
  m1 AT %QD0 : LREAL;
  m2 AT %QD2 : LREAL;
  m3 AT %QD4 : LREAL;
  m4 AT %QD6 : LREAL;
  m5 AT %QD8 : LREAL;
  m6 AT %QD10 : REAL;
  m7 AT %QD11 : LREAL;
  m8 AT %QD13 : LREAL;
  m9 AT %QD15 : LREAL;
END_VAR
  m1 := d + i;
  m2 := d * u;
  m3 := d + l;
  m4 := d + r;
  m5 := w * 1.0;
  m6 := r + 1;
  m7 := i;
  m8 := u;
  m9 := l;
END_PROGRAM

(* ---- cmp-015-lreal-multiplication-and-division.st ---- *)
PROGRAM DoubleProduct
VAR
  a : LREAL := 0.1;
  three : LREAL := 3.0;
  seven : LREAL := 7.0;
  max : LREAL := 1.7976931348623157E308;
  min : LREAL := 2.2250738585072014E-308;
  two : LREAL := 2.0;
  neg : LREAL := -1.5;
  m1 AT %QD0 : LREAL;
  m2 AT %QD2 : LREAL;
  m3 AT %QD4 : LREAL;
  m4 AT %QD6 : LREAL;
  m5 AT %QD8 : LREAL;
  d1 AT %QD10 : LREAL;
  d2 AT %QD12 : LREAL;
  d3 AT %QD14 : LREAL;
  d4 AT %QD16 : LREAL;
END_VAR
  m1 := a * three;
  m2 := neg * neg;
  m3 := max * two;
  m4 := min / two;
  m5 := min / 4503599627370496.0;
  d1 := 1.0 / three;
  d2 := a / seven;
  d3 := max / two;
  d4 := neg / two;
END_PROGRAM

(* ---- cmp-015-lreal-nan-and-infinity-propagate.st ---- *)
PROGRAM DoubleSpecials
VAR
  max : LREAL := 1.7976931348623157E308;
  one : LREAL := 1.0;
  zero : LREAL := 0.0;
  inf : LREAL;
  nan : LREAL;
  i1 AT %QD0 : LREAL;
  i2 AT %QD2 : LREAL;
  i3 AT %QD4 : LREAL;
  i4 AT %QD6 : LREAL;
  i5 AT %QD8 : LREAL;
  n1 AT %QD10 : LREAL;
  n2 AT %QD12 : LREAL;
  n3 AT %QD14 : LREAL;
  n4 AT %QD16 : LREAL;
  z1 AT %QD18 : LREAL;
END_VAR
  inf := max * 10.0;
  nan := inf - inf;
  i1 := inf;
  i2 := -inf;
  i3 := inf + one;
  i4 := one / inf;
  i5 := -one / inf;
  n1 := nan;
  n2 := nan + one;
  n3 := zero * inf;
  n4 := inf / inf;
  z1 := -zero;
END_PROGRAM

(* ---- cmp-015-lreal-narrowed-to-real-is-reported.st ---- *)
PROGRAM Narrowing
VAR
  d : LREAL := 0.1;
  r AT %QD0 : REAL;
  s AT %QD1 : REAL;
END_VAR
  r := d;
  s := d * 2.0;
END_PROGRAM

(* ---- cmp-015-lreal-transcendental-functions-compute-in-real.st ---- *)
PROGRAM DoubleLibrary
VAR
  x : LREAL := 0.5;
  ten : LREAL := 10.0;
  e1 : LREAL := 1.0;
  tol : LREAL := 0.00001;
  sin_ok AT %QX512.0 : BOOL;
  cos_ok AT %QX512.1 : BOOL;
  exp_ok AT %QX512.2 : BOOL;
  ln_ok AT %QX512.3 : BOOL;
  atan_ok AT %QX512.4 : BOOL;
  sqrt_ok AT %QX512.5 : BOOL;
END_VAR
  sin_ok := ABS(SIN(x) - 0.479425538604203) < tol;
  cos_ok := ABS(COS(x) - 0.8775825618903728) < tol;
  exp_ok := ABS(EXP(e1) - 2.718281828459045) < tol;
  ln_ok := ABS(LN(ten) - 2.302585092994046) < tol;
  atan_ok := ABS(ATAN(x) - 0.4636476090008061) < tol;
  sqrt_ok := SQRT(ten) = 3.1622776601683795;
END_PROGRAM

(* ---- cmp-015-lreal-trunc-and-round.st ---- *)
PROGRAM DoubleRounding
VAR
  a : LREAL := 2.7;
  b : LREAL := -2.7;
  h : LREAL := 2.5;
  nh : LREAL := -2.5;
  almost : LREAL := 0.49999999999999994;
  edge : LREAL := 4503599627370495.5;
  huge : LREAL := 1.0E300;
  small : LREAL := 0.3;
  t1 AT %QD0 : LREAL;
  t2 AT %QD2 : LREAL;
  t3 AT %QD4 : LREAL;
  t4 AT %QD6 : LREAL;
  r1 AT %QD8 : LREAL;
  r2 AT %QD10 : LREAL;
  r3 AT %QD12 : LREAL;
  r4 AT %QD14 : LREAL;
  r5 AT %QD16 : LREAL;
  r6 AT %QD18 : LREAL;
END_VAR
  t1 := TRUNC(a);
  t2 := TRUNC(b);
  t3 := TRUNC(huge);
  t4 := TRUNC(small);
  r1 := ROUND(h);
  r2 := ROUND(nh);
  r3 := ROUND(almost);
  r4 := ROUND(edge);
  r5 := ROUND(a);
  r6 := ROUND(huge);
END_PROGRAM

(* ---- cmp-015-lword-shifts-and-rotates-use-64-bits.st ---- *)
PROGRAM Shifts
VAR
  v : LWORD := 16#8000000000000001;
  w : LWORD := 16#0123456789ABCDEF;
  l1 AT %QD0 : LWORD;
  l2 AT %QD2 : LWORD;
  l3 AT %QD4 : LWORD;
  l4 AT %QD6 : LWORD;
  r1 AT %QD8 : LWORD;
  r2 AT %QD10 : LWORD;
  r3 AT %QD12 : LWORD;
  r4 AT %QD14 : LWORD;
  o1 AT %QD16 : LWORD;
  o2 AT %QD18 : LWORD;
  o3 AT %QD20 : LWORD;
  o4 AT %QD22 : LWORD;
  p1 AT %QD24 : LWORD;
  p2 AT %QD26 : LWORD;
  p3 AT %QD28 : LWORD;
END_VAR
  l1 := SHL(v, 1);
  l2 := SHL(w, 32);
  l3 := SHL(w, 63);
  l4 := SHL(w, 64);
  r1 := SHR(v, 1);
  r2 := SHR(w, 36);
  r3 := SHR(v, 63);
  r4 := SHR(v, 64);
  o1 := ROL(v, 1);
  o2 := ROL(w, 40);
  o3 := ROL(w, 0);
  o4 := ROL(w, 64);
  p1 := ROR(v, 1);
  p2 := ROR(w, 12);
  p3 := ROR(w, 65);
END_PROGRAM

(* ---- cmp-015-mixed-width-locals-keep-their-values.st ---- *)
PROGRAM Mixed
VAR
  flag : BOOL;
  small : SINT;
  word : INT;
  odd : BYTE;
  wide : DINT;
  ratio : REAL;
  big : LINT;
  tail : BOOL;
  o_word AT %QW0 : INT;
  o_wide AT %QD1 : DINT;
  o_ratio AT %QD2 : REAL;
  o_small AT %QB12 : SINT;
  o_odd AT %QB13 : BYTE;
  o_flag AT %QX14.0 : BOOL;
  o_tail AT %QX14.1 : BOOL;
  o_big AT %QX14.2 : BOOL;
END_VAR
  flag := TRUE;
  small := -7;
  word := -1234;
  odd := 201;
  wide := -70000;
  ratio := 2.5;
  big := 5000000000;
  tail := TRUE;
  o_word := word;
  o_wide := wide;
  o_ratio := ratio;
  o_small := small;
  o_odd := odd;
  o_flag := flag;
  o_tail := tail;
  o_big := big = 5000000000;
END_PROGRAM

(* ---- cmp-015-ulint-case-label-above-2-63.st ---- *)
PROGRAM UnsignedCase
VAR
  sel : ULINT := 18446744073709551615;
  r AT %QD0 : DINT;
END_VAR
  CASE sel OF
    0: r := 1;
    9223372036854775808..18446744073709551615: r := 2;
  ELSE r := 3;
  END_CASE;
END_PROGRAM

(* ---- cmp-015-ulint-compares-unsigned.st ---- *)
PROGRAM Unsigned
VAR
  top : ULINT := 18446744073709551615;
  mask : LWORD := 4294967296;
  all_ones : LWORD := 18446744073709551615;
  above AT %QX0.0 : BOOL;
  and_high AT %QX0.1 : BOOL;
  not_zero AT %QX0.2 : BOOL;
  xor_self AT %QX0.3 : BOOL;
END_VAR
  above := top > 1;
  and_high := (all_ones AND mask) = mask;
  not_zero := NOT mask = 18446744069414584319;
  xor_self := (all_ones XOR all_ones) = 0;
END_PROGRAM

(* ---- cmp-015-ulint-division-above-2-63.st ---- *)
PROGRAM UnsignedQuotients
VAR
  top : ULINT := 18446744073709551615;
  mid : ULINT := 9223372036854775808;
  two : ULINT := 2;
  ten : ULINT := 10;
  three : ULINT := 3;
  seven : ULINT := 7;
  q1 AT %QD0 : ULINT;
  q2 AT %QD2 : ULINT;
  q3 AT %QD4 : ULINT;
  q4 AT %QD6 : ULINT;
  r1 AT %QD8 : ULINT;
  r2 AT %QD10 : ULINT;
  r3 AT %QD12 : ULINT;
END_VAR
  q1 := top / two;
  q2 := mid / three;
  q3 := top / top;
  q4 := two / top;
  r1 := top MOD ten;
  r2 := mid MOD seven;
  r3 := top MOD mid;
END_PROGRAM

(* ---- cmp-015-ulint-division-by-zero-faults.st ---- *)
PROGRAM ByZero
VAR
  n : ULINT := 5;
  z : ULINT;
  r AT %QD0 : ULINT;
END_VAR
  r := n / z;
END_PROGRAM

(* ---- cmp-015-ulint-for-counter-up-to-the-top.st ---- *)
PROGRAM TopFor
VAR
  k : ULINT;
  hits : ULINT;
  res_hits AT %QD0 : ULINT;
  res_k AT %QD2 : ULINT;
END_VAR
  FOR k := 18446744073709551610 TO 18446744073709551613 DO
    hits := hits + 1;
  END_FOR;
  res_hits := hits;
  res_k := k;
END_PROGRAM

(* ---- cmp-015-ulint-modulo-by-zero-faults.st ---- *)
PROGRAM ByZero
VAR
  n : ULINT := 5;
  z : ULINT;
  r AT %QD0 : ULINT;
END_VAR
  r := n MOD z;
END_PROGRAM

(* ---- cmp-015-ulint-multiplication-is-unsigned.st ---- *)
PROGRAM UnsignedProduct
VAR
  big : ULINT := 18446744073709551615;
  half : ULINT := 9223372036854775808;
  t : ULINT := 3;
  w : LWORD := 16#0123456789ABCDEF;
  p1 AT %QD0 : ULINT;
  p2 AT %QD2 : ULINT;
  p3 AT %QD4 : LWORD;
  p4 AT %QD6 : ULINT;
END_VAR
  p1 := big * big;
  p2 := half * t;
  p3 := w * 16#10;
  p4 := half * 2;
END_PROGRAM

(* ---- cmp-016-dint-abs-min.st ---- *)
PROGRAM Absolute
VAR
  a : DINT := -2147483647;
  q AT %QD0 : DINT;
END_VAR
  a := a - 1;
  q := ABS(a);
END_PROGRAM

(* ---- cmp-016-dint-add-wraps.st ---- *)
PROGRAM Wrap
VAR
  a : DINT := 2147483647;
  q AT %QD0 : DINT;
END_VAR
  q := a + 1;
END_PROGRAM

(* ---- cmp-016-dint-min-divided-by-minus-one.st ---- *)
PROGRAM MinDiv
VAR
  a : DINT := -2147483647;
  m : DINT := -1;
  q AT %QD0 : DINT;
END_VAR
  a := a - 1;
  q := a / m;
END_PROGRAM

(* ---- cmp-016-dint-min-modulo-minus-one.st ---- *)
PROGRAM MinMod
VAR
  a : DINT := -2147483647;
  m : DINT := -1;
  q AT %QD0 : DINT := 5;
END_VAR
  a := a - 1;
  q := a MOD m;
END_PROGRAM

(* ---- cmp-016-dint-mul-wraps.st ---- *)
PROGRAM Wrap
VAR
  a : DINT := 100000;
  q AT %QD0 : DINT;
END_VAR
  q := a * a;
END_PROGRAM

(* ---- cmp-016-dint-negate-min.st ---- *)
PROGRAM Negate
VAR
  a : DINT := -2147483647;
  q AT %QD0 : DINT;
END_VAR
  a := a - 1;
  q := -a;
END_PROGRAM

(* ---- cmp-016-dint-sub-wraps.st ---- *)
PROGRAM Wrap
VAR
  a : DINT := -2147483647;
  q AT %QD0 : DINT;
END_VAR
  q := a - 2;
END_PROGRAM

(* ---- cmp-016-real-nan-to-dint.st ---- *)
PROGRAM NotANumber
VAR
  big : REAL := 1.0E38;
  inf : REAL;
  nan : REAL;
  q AT %QD0 : DINT := 7;
END_VAR
  inf := big * big;
  nan := inf - inf;
  q := REAL_TO_DINT(nan);
END_PROGRAM

(* ---- cmp-016-real-out-of-range-to-dint.st ---- *)
PROGRAM Saturate
VAR
  high : REAL := 3.0E9;
  low : REAL;
  q_high AT %QD0 : DINT;
  q_low AT %QD4 : DINT;
END_VAR
  low := 0.0 - high;
  q_high := REAL_TO_DINT(high);
  q_low := REAL_TO_DINT(low);
END_PROGRAM

(* ---- cmp-016-real-to-dint-truncates-toward-zero.st ---- *)
PROGRAM Truncate
VAR
  up : REAL := 1.9;
  down : REAL;
  q_up AT %QD0 : DINT;
  q_down AT %QD4 : DINT;
END_VAR
  down := 0.0 - up;
  q_up := REAL_TO_DINT(TRUNC(up));
  q_down := REAL_TO_DINT(TRUNC(down));
END_PROGRAM

(* ---- cmp-016-shift-by-the-width-or-more.st ---- *)
PROGRAM Shifts
VAR
  one : DWORD := 1;
  top : DWORD := 2147483647;
  width : DINT := 32;
  negative : DINT := -1;
  shl_width AT %QD0 : DWORD;
  shr_width AT %QD4 : DWORD;
  shl_negative AT %QD8 : DWORD;
END_VAR
  shl_width := SHL(one, width);
  shr_width := SHR(top, width);
  shl_negative := SHL(one, negative);
END_PROGRAM

(* ---- cmp-017-date-assign-and-compare.st ---- *)
PROGRAM Calendar
VAR
  first : DATE := D#2024-01-01;
  second : DATE := D#2025-06-30;
  copy : DATE;
  before AT %QX0.0 : BOOL;
  same AT %QX0.1 : BOOL;
  differ AT %QX0.2 : BOOL;
END_VAR
  copy := first;
  before := first < second;
  same := copy = D#2024-01-01;
  differ := copy <> second;
END_PROGRAM

(* ---- cmp-017-dt-compare-and-assign.st ---- *)
PROGRAM Stamp
VAR
  early : DT := DT#1970-01-01-00:00:01;
  late : DT := DT#2024-01-01-00:00:00;
  copy : DT;
  before AT %QX0.0 : BOOL;
  same AT %QX0.1 : BOOL;
END_VAR
  copy := late;
  before := early < copy;
  same := copy = DT#2024-01-01-00:00:00;
END_PROGRAM

(* ---- cmp-017-time-arithmetic-above-24-days.st ---- *)
PROGRAM Long
VAR
  a : TIME := T#30d;
  sum AT %QD0 : TIME;
  half AT %QD4 : TIME;
  bigger AT %QX8.0 : BOOL;
  smaller AT %QX8.1 : BOOL;
END_VAR
  sum := a + T#10d;
  half := a / 2;
  bigger := sum > T#35d;
  smaller := a < T#35d;
END_PROGRAM

(* ---- cmp-017-time-compare-short.st ---- *)
PROGRAM Short
VAR
  span : TIME := T#2s;
  longer AT %QX0.0 : BOOL;
END_VAR
  longer := span > T#1s;
END_PROGRAM

(* ---- cmp-017-time-compound-literal.st ---- *)
PROGRAM Duration
VAR
  t AT %QD0 : TIME;
END_VAR
  t := T#1h30m;
END_PROGRAM

(* ---- cmp-017-time-fraction-on-the-last-unit.st ---- *)
PROGRAM Parts
VAR
  a AT %QD0 : TIME;
  b AT %QD4 : TIME;
END_VAR
  a := T#1h30.5m;
  b := T#0.25s;
END_PROGRAM

(* ---- cmp-017-time-fractional-literal.st ---- *)
PROGRAM Duration
VAR
  t AT %QD0 : TIME;
END_VAR
  t := T#1.5s;
END_PROGRAM

(* ---- cmp-017-time-literal-above-the-range.st ---- *)
PROGRAM Over
VAR
  t AT %QD0 : TIME;
END_VAR
  t := T#50d;
END_PROGRAM

(* ---- cmp-017-time-literal-below-a-millisecond.st ---- *)
PROGRAM Fine
VAR
  t AT %QD0 : TIME;
END_VAR
  t := T#1.5ms;
END_PROGRAM

(* ---- cmp-017-time-literal-negative.st ---- *)
PROGRAM Negative
VAR
  t AT %QD0 : TIME;
END_VAR
  t := T#-1s;
END_PROGRAM

(* ---- cmp-017-time-literal-units-out-of-order.st ---- *)
PROGRAM Order
VAR
  t AT %QD0 : TIME;
END_VAR
  t := T#30m1h;
END_PROGRAM

(* ---- cmp-017-time-maximum-literal.st ---- *)
PROGRAM Largest
VAR
  t AT %QD0 : TIME;
END_VAR
  t := T#49d17h2m47s295ms;
END_PROGRAM

(* ---- cmp-017-time-over-24-days.st ---- *)
PROGRAM Long
VAR
  span : TIME := T#30d;
  longer AT %QX0.0 : BOOL;
END_VAR
  longer := span > T#1d;
END_PROGRAM

(* ---- cmp-017-time-subtraction-without-spaces.st ---- *)
PROGRAM Elapsed
VAR
  d AT %QD0 : TIME;
END_VAR
  d := T#5s-T#3s;
END_PROGRAM

(* ---- cmp-017-time-underscores-and-all-units.st ---- *)
PROGRAM Parts
VAR
  t AT %QD0 : TIME;
END_VAR
  t := T#1d_2h_3m_4s_5ms;
END_PROGRAM

(* ---- cmp-017-tod-compare-and-subtract-time.st ---- *)
PROGRAM Clock
VAR
  late : TOD := TOD#13:00:00;
  early : TOD := TOD#12:30:00;
  after AT %QX0.0 : BOOL;
  back AT %QX0.1 : BOOL;
  shifted AT %QD1 : TOD;
END_VAR
  after := late > early;
  shifted := late - T#30m;
  back := shifted = early;
END_PROGRAM

(* ---- cmp-017-tod-plus-time.st ---- *)
PROGRAM Clock
VAR
  start : TOD := TOD#12:30:00;
  later AT %QD0 : TOD;
END_VAR
  later := start + T#1h;
END_PROGRAM

(* ---- cmp-017-ton-with-a-30-day-preset-is-not-done.st ---- *)
PROGRAM Delay
VAR
  wait : TON;
  done AT %QX0.0 : BOOL;
END_VAR
  wait(IN := TRUE, PT := T#30d);
  done := wait.Q;
END_PROGRAM

(* ---- cmp-018-argument-does-not-fit.st ---- *)
FUNCTION Keep : SINT
VAR_INPUT
  a : SINT;
END_VAR
  Keep := a;
END_FUNCTION

PROGRAM Overflow
VAR
  x : SINT;
END_VAR
  x := Keep(300);
END_PROGRAM

(* ---- cmp-018-array-initializer-does-not-fit.st ---- *)
PROGRAM Overflow
VAR
  items : ARRAY[0..1] OF SINT := [1, 300];
END_VAR
END_PROGRAM

(* ---- cmp-018-assigned-constant-does-not-fit.st ---- *)
PROGRAM Overflow
VAR
  level : USINT;
END_VAR
  level := -1;
END_PROGRAM

(* ---- cmp-018-constant-does-not-fit.st ---- *)
PROGRAM Overflow
VAR
  small : SINT := 300;
END_VAR
  small := small + 1;
END_PROGRAM

(* ---- cmp-018-constant-expression-does-not-fit.st ---- *)
PROGRAM Overflow
VAR
  small : SINT := 100 + 100;
END_VAR
END_PROGRAM

(* ---- cmp-018-constants-at-the-limits-of-their-types.st ---- *)
PROGRAM Limits
VAR
  low : SINT := -128;
  high : SINT := 127;
  top : USINT := 255;
  wide : INT := -32768 + 65535;
  mask : BYTE := 16#FF;
  big : UDINT := 4294967295;
  out_low AT %QB0 : SINT;
  out_high AT %QB1 : SINT;
  out_top AT %QB2 : USINT;
  out_wide AT %QW2 : INT;
  out_big AT %QD2 : UDINT;
END_VAR
  out_low := low;
  out_high := high;
  out_top := top;
  out_wide := wide;
  out_big := big;
END_PROGRAM

(* ---- cmp-018-named-constant-does-not-fit.st ---- *)
PROGRAM Overflow
VAR CONSTANT
  limit : INT := 20000;
END_VAR
VAR
  doubled : INT;
END_VAR
  doubled := limit * 2;
END_PROGRAM

(* ---- cmp-019-assignment-between-different-structures-rejected.st ---- *)
TYPE Pt : STRUCT x : INT; y : INT; END_STRUCT END_TYPE
TYPE Qt : STRUCT x : INT; y : INT; END_STRUCT END_TYPE

PROGRAM Main
VAR
  p : Pt;
  q : Qt;
END_VAR
  q := p;
END_PROGRAM

(* ---- cmp-019-function-returning-a-structure-rejected.st ---- *)
TYPE Pt : STRUCT x : INT; y : INT; END_STRUCT END_TYPE

FUNCTION Make : Pt
VAR_INPUT a : INT; END_VAR
  Make.x := a;
END_FUNCTION

PROGRAM Main
VAR
  p : Pt;
END_VAR
  p := Make(1);
END_PROGRAM

(* ---- cmp-019-nested-struct-member.st ---- *)
TYPE Inner : STRUCT v : INT; END_STRUCT END_TYPE
TYPE Outer : STRUCT a : INT; inner : Inner; END_STRUCT END_TYPE

PROGRAM Nested
VAR
  o : Outer;
  seen AT %QW0 : INT;
END_VAR
  o.inner.v := 5;
  seen := o.inner.v;
END_PROGRAM

(* ---- cmp-019-nested-struct-wide-leaf.st ---- *)
TYPE Inner : STRUCT a : DINT; b : INT; END_STRUCT END_TYPE
TYPE Outer : STRUCT n : INT; inner : Inner; tail : DINT; END_STRUCT END_TYPE

PROGRAM Main
VAR
  o : Outer;
  oa AT %QD0 : DINT;
  ob AT %QW2 : INT;
  ot AT %QD2 : DINT;
  on AT %QW6 : INT;
END_VAR
  o.n := -2;
  o.inner.a := 70000;
  o.inner.b := -300;
  o.tail := 80000;
  oa := o.inner.a;
  ob := o.inner.b;
  ot := o.tail;
  on := o.n;
END_PROGRAM

(* ---- cmp-019-struct-as-parameter.st ---- *)
TYPE Pt : STRUCT x : INT; y : INT; z : DINT; END_STRUCT END_TYPE

FUNCTION SumXY : INT
VAR_INPUT p : Pt; END_VAR
  SumXY := p.x + p.y;
END_FUNCTION

PROGRAM Param
VAR
  point : Pt;
  total AT %QW0 : INT;
END_VAR
  point.x := 3;
  point.y := 4;
  total := SumXY(point);
END_PROGRAM

(* ---- cmp-019-struct-assignment-copies-all.st ---- *)
TYPE Pt : STRUCT x : INT; y : INT; z : DINT; END_STRUCT END_TYPE

PROGRAM Copy
VAR
  p : Pt;
  q : Pt;
  seen AT %QD0 : DINT;
END_VAR
  p.x := 1;
  p.z := 7;
  q := p;
  seen := q.z;
END_PROGRAM

(* ---- cmp-019-struct-assignment-nested.st ---- *)
TYPE Inner : STRUCT a : DINT; b : INT; END_STRUCT END_TYPE
TYPE Outer : STRUCT n : INT; inner : Inner; tail : DINT; END_STRUCT END_TYPE

PROGRAM Main
VAR
  src : Outer;
  dst : Outer;
  oa AT %QD0 : DINT;
  ot AT %QD1 : DINT;
  on AT %QW4 : INT;
END_VAR
  src.n := 5;
  src.inner.a := 70000;
  src.tail := 80000;
  dst := src;
  src.inner.a := 1;
  src.tail := 2;
  oa := dst.inner.a;
  ot := dst.tail;
  on := dst.n;
END_PROGRAM

(* ---- cmp-019-struct-dint-member.st ---- *)
TYPE Pt : STRUCT x : INT; y : INT; z : DINT; END_STRUCT END_TYPE

PROGRAM Member
VAR
  p : Pt;
  seen AT %QD0 : DINT;
END_VAR
  p.z := 100000;
  seen := p.z;
END_PROGRAM

(* ---- cmp-019-struct-initialiser-defaults.st ---- *)
TYPE Pt : STRUCT x : INT := 7; y : INT := 8; z : DINT := 100000; END_STRUCT END_TYPE

PROGRAM Main
VAR
  p : Pt := (y := 20);
  q : Pt;
  px AT %QW0 : INT;
  py AT %QW1 : INT;
  pz AT %QD1 : DINT;
  qx AT %QW4 : INT;
END_VAR
  px := p.x;
  py := p.y;
  pz := p.z;
  qx := q.x;
END_PROGRAM

(* ---- cmp-019-struct-initialiser.st ---- *)
TYPE Pt : STRUCT x : INT; y : INT; z : DINT; END_STRUCT END_TYPE

PROGRAM Init
VAR
  p : Pt := (x := 1, y := 2);
  seen AT %QW0 : INT;
END_VAR
  seen := p.y;
END_PROGRAM

(* ---- cmp-019-struct-int-member.st ---- *)
TYPE Pt : STRUCT x : INT; y : INT; z : DINT; END_STRUCT END_TYPE

PROGRAM Member
VAR
  p : Pt;
  seen AT %QW0 : INT;
END_VAR
  p.x := 1000;
  seen := p.x;
END_PROGRAM

(* ---- cmp-019-struct-members-do-not-overlap.st ---- *)
TYPE Mixed : STRUCT f : BOOL; b : BYTE; i : INT; d : DINT; r : REAL; END_STRUCT END_TYPE

PROGRAM Main
VAR
  m : Mixed;
  oflag AT %QX0.0 : BOOL;
  ob AT %QB1 : BYTE;
  oi AT %QW1 : INT;
  od AT %QD1 : DINT;
  orr AT %QD2 : REAL;
END_VAR
  m.d := 123456;
  m.r := 0.5;
  m.i := 31000;
  m.b := 250;
  m.f := TRUE;
  oflag := m.f;
  ob := m.b;
  oi := m.i;
  od := m.d;
  orr := m.r;
END_PROGRAM

(* ---- cmp-019-struct-negative-members.st ---- *)
TYPE Pt : STRUCT a : SINT; b : INT; c : DINT; END_STRUCT END_TYPE

PROGRAM Main
VAR
  p : Pt;
  sa AT %QB0 : SINT;
  sb AT %QW1 : INT;
  sc AT %QD1 : DINT;
END_VAR
  p.a := -5;
  p.b := -1000;
  p.c := -100000;
  sa := p.a;
  sb := p.b;
  sc := p.c;
END_PROGRAM

(* ---- cmp-019-struct-parameter-keeps-every-member.st ---- *)
TYPE Pt : STRUCT x : INT; y : INT; z : DINT; END_STRUCT END_TYPE

FUNCTION Tail : DINT
VAR_INPUT whole : Pt; END_VAR
  Tail := whole.z;
END_FUNCTION

FUNCTION Bump : INT
VAR_INPUT copy : Pt; END_VAR
  copy.x := 99;
  Bump := copy.x;
END_FUNCTION

PROGRAM Main
VAR
  point : Pt;
  z AT %QD0 : DINT;
  bumped AT %QW2 : INT;
  kept AT %QW3 : INT;
END_VAR
  point.x := 3;
  point.z := 100000;
  z := Tail(point);
  bumped := Bump(point);
  kept := point.x;
END_PROGRAM

(* ---- cmp-019-struct-small-members.st ---- *)
TYPE Pt : STRUCT x : INT; y : INT; z : DINT; END_STRUCT END_TYPE

PROGRAM Member
VAR
  p : Pt;
  total AT %QW0 : INT;
END_VAR
  p.x := 3;
  p.y := 4;
  total := p.x + p.y;
END_PROGRAM

(* ---- cmp-019-structure-as-a-number-rejected.st ---- *)
TYPE Pt : STRUCT x : INT; y : INT; END_STRUCT END_TYPE

PROGRAM Main
VAR
  p : Pt;
  n : DINT;
END_VAR
  n := p;
END_PROGRAM

(* ---- cmp-020-enum-array.st ---- *)
TYPE St : (IDLE, RUN, FAULT); END_TYPE

PROGRAM Main
VAR
  a : ARRAY[0..2] OF St;
  one AT %QW0 : INT;
  two AT %QW1 : INT;
  zero AT %QW2 : INT;
END_VAR
  a[1] := RUN;
  a[2] := FAULT;
  one := a[1];
  two := a[2];
  zero := a[0];
END_PROGRAM

(* ---- cmp-020-enum-case-labels.st ---- *)
TYPE St : (IDLE, RUN, FAULT := 5); END_TYPE

PROGRAM Main
VAR
  s : St;
  r AT %QW0 : INT;
END_VAR
  s := St#FAULT;
  CASE s OF
    IDLE: r := 10;
    RUN: r := 20;
    FAULT: r := 50;
  END_CASE;
END_PROGRAM

(* ---- cmp-020-enum-compare-ignores-neighbour.st ---- *)
TYPE St : (IDLE, RUN); END_TYPE

PROGRAM Machine
VAR
  state : St;
  next : INT;
  running AT %QX0.0 : BOOL;
END_VAR
  state := RUN;
  next := 7;
  running := state = RUN;
END_PROGRAM

(* ---- cmp-020-enum-members-keep-neighbours.st ---- *)
TYPE St : (IDLE, RUN, FAULT); END_TYPE
TYPE Machine : STRUCT before : INT; state : St; after : DINT; END_STRUCT END_TYPE

PROGRAM Main
VAR
  m : Machine;
  ob AT %QW0 : INT;
  os AT %QW1 : INT;
  oa AT %QD1 : DINT;
END_VAR
  m.before := 11;
  m.after := 222222;
  m.state := FAULT;
  ob := m.before;
  os := m.state;
  oa := m.after;
END_PROGRAM

(* ---- cmp-020-enum-qualified-case-label.st ---- *)
TYPE St : (IDLE, RUN, FAULT); END_TYPE

PROGRAM Main
VAR
  s : St := St#RUN;
  r AT %QW0 : INT;
END_VAR
  CASE s OF
    St#IDLE: r := 10;
    St#RUN: r := 20;
    St#FAULT: r := 30;
  END_CASE;
END_PROGRAM

(* ---- cmp-020-enum-qualified-literal.st ---- *)
TYPE St : (IDLE, RUN); END_TYPE

PROGRAM Machine
VAR
  state : St;
  running AT %QX0.0 : BOOL;
END_VAR
  state := St#RUN;
  running := state = RUN;
END_PROGRAM

(* ---- cmp-020-enum-store-keeps-neighbour.st ---- *)
TYPE St : (IDLE, RUN); END_TYPE

PROGRAM Machine
VAR
  state : St;
  next : INT;
  seen AT %QW0 : INT;
END_VAR
  next := 7;
  state := RUN;
  seen := next;
END_PROGRAM
